      L     #Enc;
      T     #Data.Fall_Pos;
      L     #Data.Time_ms;
      T     #Data.Fall_ms;
      SET   ;
      S     #Data.Low;

S020: NOP   0;
NETWORK
TITLE =OFF Longer than Gap_Min = Real Gap - Close Packet

      A     #RUN;
      AN    #Sensor;
      A     #Data.Open;
      A     #Data.Low;
      JCN   S030;

      L     #Enc;
      L     #Data.Fall_Pos;
      -D    ;
      T     #D;
      L     L#0;
      >=D   ;
      JC    S031;

      L     #D;
      NEGD  ;
      T     #D;

S031: L     #D;
      L     #Gap_Min_Pulse;
      >=D   ;
      =     #CLOSE;

S030: NOP   0;
NETWORK
TITLE =Transfer End - Close Last Packet / Discard Covered One
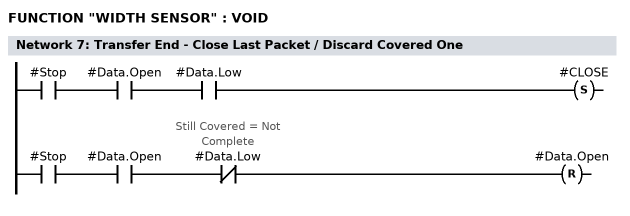

      A     #Stop;
      A     #Data.Open;
      A     #Data.Low;
      S     #CLOSE;
//;
      A     #Stop;
      A     #Data.Open;
      AN    #Data.Low; // Still Covered = Not Complete
      R     #Data.Open;

NETWORK
TITLE =Close Packet - Record Width

      A     #CLOSE;
      JCN   S090;

      A     #Data.Skip; // Partial Packet - Not Recorded
      JCN   S041;

      L     #Data.Skipped;
      L     1;
      +I    ;
      T     #Data.Skipped;
      JU    S049;

S041: L     #Data.Fall_Pos;
      L     #Data.Start_Pos;
      -D    ;
      T     #D;
      L     L#0;
      >=D   ;
      JC    S042;

      L     #D;
      NEGD  ;
      T     #D;

S042: L     #D;
      DTR   ;
      L     3.100000e-001;
      *R    ;
      RND   ;
      T     #MM;
      T     #Data.Last_Width_mm;
      L     #Data.Count;
      L     1;
      +I    ;
      T     #Data.Count;
      L     #MM;
      ITD   ;
      L     #Data.Width_Sum_mm;
      +D    ;
      T     #Data.Width_Sum_mm;
      L     #MM;
      L     #Data.Width_Min_mm;
      <I    ;
      JCN   S043;

      L     #MM;
      T     #Data.Width_Min_mm;

S043: L     #MM;
      L     #Data.Width_Max_mm;
      >I    ;
      JCN   S044;

      L     #MM;
      T     #Data.Width_Max_mm;

S044: L     #Data.Width_Sum_mm;
      L     #Data.Count;
      ITD   ;
      /D    ;
      T     #Data.Width_Avg_mm;
//;
      L     #Data.Fall_ms; // Width [mS] = Front -> End
      T     #Data.Last_Width_ms;
      L     #Data.Width_Sum_ms;
      +D    ;
      T     #Data.Width_Sum_ms;
      L     #Data.Count;
      ITD   ;
      /D    ;
      T     #Data.Width_Avg_ms;

S049: SET   ;
      R     #Data.Open;
      R     #Data.Low;
      R     #Data.Skip;

S090: NOP   0;
NETWORK
TITLE =Sensor State for Next Scan

      A     #Sensor;
      =     #Data.Was_On;
END_FUNCTION

FUNCTION "PACKET BLANKING" : VOID
TITLE =Packet Blanking - One Sensor (Shadow)
//v0.1 2026-11-19: one count per packet from a raw sensor, with the packet time
//measured at C10 (DB30 Width_ms_31, same speed on C11/C12/C21/C22).
//- Front (OFF->ON) counts if the belt has run >= Blank_Pct of a packet time
//  since the last count; an earlier front = sag of a U-Shape -> ignored.
//- Sensor still ON after Butt_Pct of a packet time = butted packet -> +1.
//- Time only runs while the belt runs (Run): a stop does not open the window.
//- Pulse: Pulse_ms long per counted packet (for FC8 later).
VERSION : 0.1


VAR_INPUT
  Sensor : BOOL ;	//Raw Packet Sensor
  Run : BOOL ;	//Belt Under the Sensor Runs
  Width_ms : INT ;	//Packet Time [mS]
  Blank_Pct : INT ;	//Blanking [%]
  Butt_Pct : INT ;	//Butted [%]
  Pulse_Len : INT ;	//Pulse [mS]
  Scan_mS : INT ;	//PLC Scan [mS]
END_VAR
VAR_OUTPUT
  Pulse : BOOL ;	//One Pulse per Counted Packet
END_VAR
VAR_IN_OUT
  D : "Blanking Struct";
END_VAR
VAR_TEMP
  BLANK : DINT ;
  BUTT : DINT ;
  CNT : BOOL ;
  BTD : BOOL ;
END_VAR
BEGIN
NETWORK
TITLE =Belt Run Time Since Last Count

      CLR   ;
      =     #CNT;
      =     #BTD;
//;
      A     #Run;
      JCN   B001;

      L     #D.T_ms;
      L     #Scan_mS;
      ITD   ;
      +D    ;
      T     #D.T_ms;
      L     #D.T_ms;
      L     L#60000;
      >D    ; // Clamp 60s
      JCN   B001;

      L     L#60000;
      T     #D.T_ms;

B001: NOP   0;
NETWORK
TITLE =Windows [mS]

      L     #Width_ms;
      ITD   ;
      L     #Blank_Pct;
      ITD   ;
      *D    ;
      L     L#100;
      /D    ;
      T     #BLANK;
//;
      L     #Width_ms;
      ITD   ;
      L     #Butt_Pct;
      ITD   ;
      *D    ;
      L     L#100;
      /D    ;
      T     #BUTT;
NETWORK
TITLE =Front - Count, or Ignore Inside Blanking (Sag)

      A     #Sensor;
      AN    #D.Was_On;
      JCN   B010;

      L     #D.Raw;
      L     1;
      +I    ;
      T     #D.Raw;
//;
      L     #D.T_ms;
      L     #BLANK;
      >=D   ;
      =     #CNT; // Front Counts
      JC    B010;

      L     #D.Sag; // Front Inside Blanking = Sag
      L     1;
      +I    ;
      T     #D.Sag;

B010: NOP   0;
NETWORK
TITLE =Sensor Still ON - Butted Packet

      A     #Sensor;
      A     #Run;
      AN    #CNT;
      JCN   B020;

      L     #D.T_ms;
      L     #BUTT;
      >=D   ;
      JCN   B020;

      L     #D.Butt;
      L     1;
      +I    ;
      T     #D.Butt;
      SET   ;
      =     #CNT;
      =     #BTD; // Next Butted Packet One Packet Time Later

B020: NOP   0;
NETWORK
TITLE =Count + Pulse

      A     #CNT;
      JCN   B030;

      L     #D.Count;
      L     1;
      +I    ;
      T     #D.Count;
      L     L#0;
      T     #D.T_ms;
      A     #BTD;
      JCN   B032;

      L     #BUTT; // Butted: T = Butt - Packet Time
      L     #Width_ms;
      ITD   ;
      -D    ;
      T     #D.T_ms;

B032: L     #Pulse_Len;
      T     #D.Pulse_ms;

B030: L     #D.Pulse_ms;
      L     0;
      >I    ;
      =     #Pulse;
      =     #D.Pulse;
      JCN   B031;

      L     #D.Pulse_ms;
      L     #Scan_mS;
      -I    ;
      T     #D.Pulse_ms;

B031: A     #Sensor;
      =     #D.Was_On;
END_FUNCTION

FUNCTION "PACKET POSITIONING" : VOID
TITLE =Packet Positioning - Flipper C7 + Pusher 2 C9 - Stop Time per Lengt
//v1.0 2026-11-23: called by FC942 v1.0. Picks the stop time of the length class
//of the packets (C4 measurement), lights the class lamp, and lets the operator
//change that class time with the HMI arrows (+/- Step_ms, Min_ms...Max_ms).
//Writes only DB15 "PACKET POSITION DB". Empty table = Default_ms = 1.5 s as before.
//v1.1 2026-11-24: HMI packet drawing: length (DBW86) + width class bits (DBX90.x).
//v1.2 2026-11-24: renumbered FC1221 -> FC1215 (same name "FLIPPER POS ADJ", no
//code change). FC942 calls it by name.
//v1.3 2026-11-24: renamed "PACKET POSITIONING". + C9 Pusher 2 conveyor: same
//length class, own table / arrows, default = "HMI_DB".CONV_9_POS_mS x 10 (as
//before). Output C9_Stop_S5T for FC950 v1.0 Timer 62.
//v1.4 2026-11-24: C9 HMI drawing: C9_Pos_Bits (one of 16 lateral positions).
//v1.5 2026-11-24: DB15 symbol renamed "PACKET POSITION DB" - no code change.
VERSION : 1.5


VAR_TEMP
  CLASS : INT ;
  T_TAB : INT ;
  T_NEW : INT ;
  T_DEF : INT ;
  T_TIME : TIME ;
  S5 : S5TIME ;
END_VAR
BEGIN
NETWORK
TITLE =Packet Length -> Class (15 mm Steps from 510 mm, 0...31)

      L     "HOUSE_KEEPING DB".C4_Packet_Length_mm;
      T     "PACKET POSITION DB".Length_mm;
      L     510;
      -I    ;
      L     15;
      /I    ;
      T     #CLASS;
      L     0;
      >=I   ;
      JC    K001;

      L     0;
      T     #CLASS;

K001: L     #CLASS;
      L     31;
      <=I   ;
      JC    K002;

      L     31;
      T     #CLASS;

K002: L     #CLASS;
      T     "PACKET POSITION DB".Class;
//;
      L     #CLASS; // Class Lamp: Bit = Class
      L     L#1;
      SLD   ;
      T     "PACKET POSITION DB".Class_Lamps;
NETWORK
TITLE =C7 Flipper - Read the Class Time (Time_ms[Class], DB15.DBW22 + 2 x

      L     #CLASS;
      SLW   1;
      L     22;
      +I    ;
      SLD   3;
      LAR1  ;
      OPN   "PACKET POSITION DB";
      L     DBW [AR1,P#0.0];
      T     #T_TAB;
NETWORK
TITLE =C7 Flipper - HMI Arrows / Reset - Change This Class Time
//The HMI sets Plus_PB / Minus_PB / Reset_PB, the PLC resets them after use:
//one press = one step.
      L     #T_TAB; // Start From the Time Used (0 = Default)
      L     0;
      <>I   ;
      JC    K010;

      L     "PACKET POSITION DB".Default_ms;
      JU    K011;

K010: L     #T_TAB;
K011: T     #T_NEW;
//;
      A     "PACKET POSITION DB".Plus_PB;
      JCN   K012;

      L     #T_NEW;
      L     "PACKET POSITION DB".Step_ms;
      +I    ;
      T     #T_NEW;

K012: A     "PACKET POSITION DB".Minus_PB;
      JCN   K013;

      L     #T_NEW;
      L     "PACKET POSITION DB".Step_ms;
      -I    ;
      T     #T_NEW;

K013: L     #T_NEW; // Clamp Min...Max
      L     "PACKET POSITION DB".Min_ms;
      >=I   ;
      JC    K014;

      L     "PACKET POSITION DB".Min_ms;
      T     #T_NEW;

K014: L     #T_NEW;
      L     "PACKET POSITION DB".Max_ms;
      <=I   ;
      JC    K015;

      L     "PACKET POSITION DB".Max_ms;
      T     #T_NEW;

K015: NOP   0;
NETWORK
TITLE =C7 Flipper - Write Back After an Arrow / Reset

      A     "PACKET POSITION DB".Reset_PB;
      JCN   K020;

      L     0; // Class Back to Default
      T     #T_TAB;
      JU    K021;

K020: A(    ;
      O     "PACKET POSITION DB".Plus_PB;
      O     "PACKET POSITION DB".Minus_PB;
      )     ;
      JCN   K022;

      L     #T_NEW;
      T     #T_TAB;

K021: L     #CLASS;
      SLW   1;
      L     22;
      +I    ;
      SLD   3;
      LAR1  ;
      OPN   "PACKET POSITION DB";
      L     #T_TAB;
      T     DBW [AR1,P#0.0];

K022: SET   ; // Momentary: Reset by the PLC
      R     "PACKET POSITION DB".Plus_PB;
      R     "PACKET POSITION DB".Minus_PB;
      R     "PACKET POSITION DB".Reset_PB;
NETWORK
TITLE =HMI Packet Drawing - Length + Width Class (4 Pairs of Level Meters)
//Width = C10 measured width (DB30 Width_mm_Cal, last verified, same order).
//0 (not measured yet) = smallest class.
      L     "PACKET POSITION DB".Length_mm;
      T     "PACKET POSITION DB".Disp_Length_mm;
//;
      L     "PACKET WIDTH DB".Width_mm_Cal;
      T     "PACKET POSITION DB".Width_mm;
//;
      L     "PACKET POSITION DB".Width_mm;
      L     "PACKET POSITION DB".Width_Lim_1;
      <I    ;
      =     "PACKET POSITION DB".Width_Class_1;
//;
      A(    ;
      L     "PACKET POSITION DB".Width_mm;
      L     "PACKET POSITION DB".Width_Lim_1;
      >=I   ;
      )     ;
      A(    ;
      L     "PACKET POSITION DB".Width_mm;
      L     "PACKET POSITION DB".Width_Lim_2;
      <I    ;
      )     ;
      =     "PACKET POSITION DB".Width_Class_2;
//;
      A(    ;
      L     "PACKET POSITION DB".Width_mm;
      L     "PACKET POSITION DB".Width_Lim_2;
      >=I   ;
      )     ;
      A(    ;
      L     "PACKET POSITION DB".Width_mm;
      L     "PACKET POSITION DB".Width_Lim_3;
      <I    ;
      )     ;
      =     "PACKET POSITION DB".Width_Class_3;
//;
      L     "PACKET POSITION DB".Width_mm;
      L     "PACKET POSITION DB".Width_Lim_3;
      >=I   ;
      =     "PACKET POSITION DB".Width_Class_4;
NETWORK
TITLE =C7 Flipper - Stop Time Used -> S5TIME for FC942 Timer 42

      L     #T_TAB;
      L     0;
      <>I   ;
      A     "PACKET POSITION DB".Use_Table;
      JC    K030;

      L     "PACKET POSITION DB".Default_ms;
      JU    K031;

K030: L     #T_TAB;
K031: T     "PACKET POSITION DB".Time_Used_ms;
      ITD   ;
      T     #T_TIME;

      CALL "TIM_S5TI" (
           IN                       := #T_TIME,
           RET_VAL                  := #S5);

      L     #S5;
      T     "PACKET POSITION DB".Stop_S5T;
NETWORK
TITLE =C9 Pusher 2 - Read the Class Time (C9_Time_ms[Class], DB15.DBW108 +

      L     "PACKET POSITION DB".Class;
      T     #CLASS;
      SLW   1;
      L     108;
      +I    ;
      SLD   3;
      LAR1  ;
      OPN   "PACKET POSITION DB";
      L     DBW [AR1,P#0.0];
      T     #T_TAB;
//;
      L     "HMI_DB".CONV_9_POS_mS; // C9 Default = HMI Time x 10 mS (as Before)
      L     10;
      *I    ;
      T     #T_DEF;
NETWORK
TITLE =C9 Pusher 2 - HMI Arrows / Reset - Change This Class Time

      L     #T_TAB;
      L     0;
      <>I   ;
      JC    C010;

      L     #T_DEF;
      JU    C011;

C010: L     #T_TAB;
C011: T     #T_NEW;
//;
      A     "PACKET POSITION DB".C9_Plus_PB;
      JCN   C012;

      L     #T_NEW;
      L     "PACKET POSITION DB".Step_ms;
      +I    ;
      T     #T_NEW;

C012: A     "PACKET POSITION DB".C9_Minus_PB;
      JCN   C013;

      L     #T_NEW;
      L     "PACKET POSITION DB".Step_ms;
      -I    ;
      T     #T_NEW;

C013: L     #T_NEW; // Clamp 1...Max (0 Means Default)
      L     1;
      >=I   ;
      JC    C014;

      L     1;
      T     #T_NEW;

C014: L     #T_NEW;
      L     "PACKET POSITION DB".Max_ms;
      <=I   ;
      JC    C015;

      L     "PACKET POSITION DB".Max_ms;
      T     #T_NEW;

C015: NOP   0;
NETWORK
TITLE =C9 Pusher 2 - Write Back After an Arrow / Reset

      A     "PACKET POSITION DB".C9_Reset_PB;
      JCN   C020;

      L     0; // Class Back to Default
      T     #T_TAB;
      JU    C021;

C020: A(    ;
      O     "PACKET POSITION DB".C9_Plus_PB;
      O     "PACKET POSITION DB".C9_Minus_PB;
      )     ;
      JCN   C022;

      L     #T_NEW;
      T     #T_TAB;

C021: L     #CLASS;
      SLW   1;
      L     108;
      +I    ;
      SLD   3;
      LAR1  ;
      OPN   "PACKET POSITION DB";
      L     #T_TAB;
      T     DBW [AR1,P#0.0];

C022: SET   ; // Momentary: Reset by the PLC
      R     "PACKET POSITION DB".C9_Plus_PB;
      R     "PACKET POSITION DB".C9_Minus_PB;
      R     "PACKET POSITION DB".C9_Reset_PB;
NETWORK
TITLE =C9 Pusher 2 - Stop Time Used -> S5TIME for FC950 Timer 62

      L     #T_TAB;
      L     0;
      <>I   ;
      A     "PACKET POSITION DB".C9_Use_Table;
      JC    C030;

      L     #T_DEF;
      JU    C031;

C030: L     #T_TAB;
C031: T     "PACKET POSITION DB".C9_Time_Used_ms;
      ITD   ;
      T     #T_TIME;

      CALL "TIM_S5TI" (
           IN                       := #T_TIME,
           RET_VAL                  := #S5);

      L     #S5;
      T     "PACKET POSITION DB".C9_Stop_S5T;
NETWORK
TITLE =C9 Pusher 2 - HMI Drawing: 1 of 16 Lateral Positions (Longer Time =

      L     "PACKET POSITION DB".C9_View_Step_ms; // Step 0 -> Copy 0
      L     0;
      >I    ;
      JC    C040;

      L     0;
      JU    C042;

C040: L     "PACKET POSITION DB".C9_Time_Used_ms;
      L     "PACKET POSITION DB".C9_View_Min_ms;
      -I    ;
      L     "PACKET POSITION DB".C9_View_Step_ms;
      /I    ;
      T     #T_NEW;
      L     0;
      >=I   ;
      JC    C041;

      L     0;
      T     #T_NEW;

C041: L     #T_NEW;
      L     15;
      <=I   ;
      L     #T_NEW;
      JC    C042;

      L     15;
C042: T     "PACKET POSITION DB".C9_Pos_Step;
//;
      L     "PACKET POSITION DB".C9_Pos_Step; // One Bit = Step
      L     L#1;
      SLD   ;
      T     "PACKET POSITION DB".C9_Pos_Bits;
END_FUNCTION

FUNCTION "LAUER CALL" : VOID
TITLE =Lauer Call
// TEXT ORG
NAME : TEXTORG
VERSION : 0.0

BEGIN
NETWORK
TITLE =

      OPN   "DB LAUER";

NETWORK
TITLE =Reset & Preset
//When the communication/control byte is in a neutral state, and those two
//internal flags are off, the FC restores default preset values in the Lauer DB.
      A(    ;
      L     "MB 150";
      L     W#16#FFF7;
      AW    ;
      L     W#16#0;
      )     ;
      ==I   ;
      AN    "M 151.6";
      AN    "M 151.7";
      JC    M001;
      JU    M002;

M001: L     2#0;
      T     DBW   76;
//;
      L     2#111100000000;
      T     DBW   72;
//;
      L     2#11100000000001;
      T     DBW   74;
//;
      L     W#16#0;
      T     DBW   32;

M002: NOP   0;
NETWORK
TITLE =
//transfer keypad/page/request words
//avoid repeated copying every scan
//only copy
//once per trigger edge/state
      A     "M 0.3";
      AN    "M 200.0";
      JC    M003;
      A     "M 0.2";
      AN    "M 200.1";
      JC    M004;
      JU    M005;

M003: L     "MW 150";
      T     "MW 118";
//;
      L     "MW 152";
      T     "MW 120";
//;
      A     "M 0.3";
      S     "M 200.0";
      R     "M 200.1";
      JU    M005;

M004: L     "MW 118";
      T     "MW 150";
//;
      L     "MW 120";
      T     "MW 152";
//;
      A     "M 0.2";
      S     "M 200.1";
      R     "M 200.0";

M005: NOP   0;
NETWORK
TITLE =
//reopen "DB LAUER"
//
//load DBW48
//
//call LAUER KEYS 1
      OPN   "DB LAUER";
      L     DBW   48;
      CALL "LAUER KEYS 1" ;
NETWORK
TITLE =

      CALL "LAUER SERVICE" ;

NETWORK
TITLE =

      CALL "LAUER KEYS 2" ;

NETWORK
TITLE =

      CALL "LAUER KEYS 3" ;

NETWORK
TITLE =

      CALL "LAUER MESSAGE1" ;

NETWORK
TITLE =

//      CALL  "LAUER"

NETWORK
TITLE =

      CALL "LAUER MESSAGE2" ;

END_FUNCTION

FUNCTION "SETUP" : VOID
TITLE =Setup Values
//Do Not Change These Values !!!
NAME : SETUP
VERSION : 0.1

BEGIN
NETWORK
TITLE =Setup Values - Slat Conveyor 3

      L     8000;
      T     "COLLATORS DB".Conveyor_Length_C3;
NETWORK
TITLE =Setup Values - Conveyor 4

      L     800; //900
      T     "COLLATORS DB".Surface_Length_C4;
NETWORK
TITLE =Setup Value  - TurnTable - Need " Packet IN " to Start

      S     "M 47.4";

NETWORK
TITLE =Setup Values - Conveyor 10

      L     13000;
      T     "COLLATORS DB".Surface_Length_10;
NETWORK
TITLE =Counter Setup


      S     "M 167.7";
NETWORK
TITLE =Packet Counter Constants 11.0 & 5.5

      L     1.000000e+001;
      T     "DB UTILITY".LENGTH_CONST;
//;
      L     5.200000e-001;
      T     "DB UTILITY".WIDTH_CONST;
NETWORK
TITLE =HMI - Conveyor Time

      L     150;
      T     "HMI_DB".CONV_7_POS_mS;
//;
      L     30;
      T     "HMI_DB".CONV_8_POS_FWD_mS;
//;
      L     70;
      T     "HMI_DB".CONV_8_POS_REV_mS;
//;
      L     15;
      T     "HMI_DB".CONV_9_POS_mS;
NETWORK
TITLE =HMI Control - Reset

      R     "HMI_DB".SERVICE_SW_1_STATUS;
      R     "HMI_DB".SERVICE_SW_2_STATUS;
      R     "HMI_DB".SERVICE_SW_3_STATUS;
      R     "HMI_DB".SERVICE_SW_1_2_STATUS;
END_FUNCTION

FUNCTION "SENSOR DE-BOUNCER" : VOID
TITLE =Sensor Debouncer
//Counting Foul Sensor Switching of less than PreSet Time
VERSION : 0.2


VAR_INPUT
  Bit_0 : BOOL ;
  Bit_1 : BOOL ;
  Preset_mS : INT ;
  Debounce_mS : INT ;
  Plc_Scan_mS : INT ;
END_VAR
VAR_IN_OUT
  Rising_Pulse_1 : BOOL ;	//Db Struct
  Rising_Pulse_2 : BOOL ;	//Db Struct
  Rising_Pulse_3 : BOOL ;	//Db Struct
  Rising_Pulse_4 : BOOL ;	//Db Struct
  Rising_Pulse_5 : BOOL ;	//Db Struct
  Rising_Pulse_6 : BOOL ;	//Db Struct
  Rising_Pulse_7 : BOOL ;	//Db Struct
  Rising_Pulse_8 : BOOL ;	//Db Struct
  Memory_Bit_1 : BOOL ;	//Db Struct
  Memory_Bit_2 : BOOL ;	//Db Struct
  Memory_Bit_3 : BOOL ;	//Db Struct
  Memory_Bit_4 : BOOL ;	//Db Struct
  Memory_Bit_5 : BOOL ;	//Db Struct
  Memory_Bit_6 : BOOL ;	//Db Struct
  Spare_1 : BOOL ;	//Db Struct
  Spare_2 : BOOL ;	//Db Struct
  Word_Buffer_1 : INT ;	//Db Struct
  Word_Buffer_2 : INT ;	//Db Struct
  Word_Result : INT ;	//Db Struct
  Word_Count_Limit : INT ;	//Db Data
  Word_Count : INT ;	//Db/HMI Data
END_VAR
VAR_TEMP
  MEMORY_1 : BOOL ;
  MEMORY_2 : BOOL ;
  MEMORY_3 : BOOL ;
END_VAR
BEGIN
NETWORK
TITLE =Init on First Call

      A     #Memory_Bit_6;
      JNB   INI1;
      JU    INI2;

INI1: L     0;
      T     #Word_Buffer_1;
      T     #Word_Buffer_2;
      R     #Memory_Bit_1;
      R     #Memory_Bit_2;
      R     #Memory_Bit_3;
      R     #Memory_Bit_4;
      R     #Memory_Bit_5;
      S     #Memory_Bit_6;

INI2: NOP   0;

NETWORK
TITLE =Input Bits - Start Event
//- #Bit_0 : Conveyor X InFeed Sensor
//- #Bit_1 : Conveyor X Exit Sensor
      A     #Bit_0;
      FP    #Rising_Pulse_1;
      JNB   K001;
      L     0;
      T     #Word_Buffer_1;
      R     #Memory_Bit_4;
      S     #Memory_Bit_1;

K001: NOP   0;

      A     #Bit_1;
      FP    #Rising_Pulse_2;
      JNB   K002;
      L     0;
      T     #Word_Buffer_2;
      S     #Memory_Bit_2;

K002: NOP   0;

NETWORK
TITLE =TimeBase
//TimeBase -> ScanTime
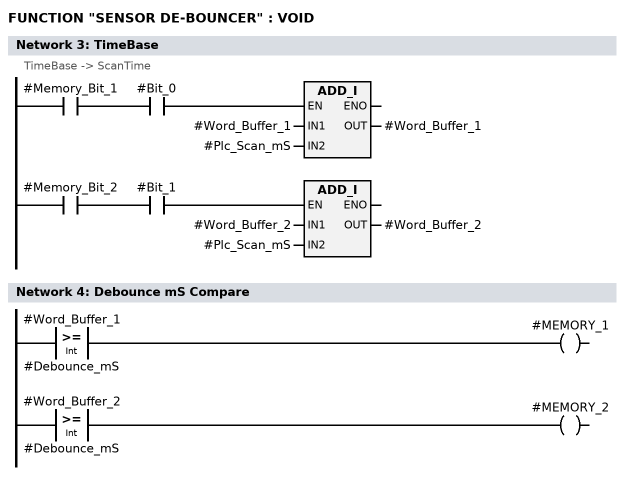
      A     #Memory_Bit_1;
      A     #Bit_0;
      JNB   K003;
      L     #Word_Buffer_1;
      L     #Plc_Scan_mS;
      +I    ;
      T     #Word_Buffer_1;

K003: NOP   0;

      A     #Memory_Bit_2;
      A     #Bit_1;
      JNB   K004;
      L     #Word_Buffer_2;
      L     #Plc_Scan_mS;
      +I    ;
      T     #Word_Buffer_2;

K004: NOP   0;

NETWORK
TITLE =Debounce mS Compare

      A(    ;
      L     #Word_Buffer_1;
      L     #Debounce_mS;
      >=I   ;
      )     ;
      =     #MEMORY_1;
//;
      A(    ;
      L     #Word_Buffer_2;
      L     #Debounce_mS;
      >=I   ;
      )     ;
      =     #MEMORY_2;

NETWORK
TITLE =Add to Packet Number with Bit_0
//Validated ON event on Bit_0 adds +1 one time
      A     #Memory_Bit_1;
      A     #MEMORY_1;
      A     #Bit_0;
      FP    #Rising_Pulse_4;
      JNB   K005;
      L     #Word_Count;
      L     1;
      +I    ;
      T     #Word_Count;
      R     #Memory_Bit_1;

K005: NOP   0;

NETWORK
TITLE =Subtract from Packet Number with Bit_1
//Validated ON event on Bit_1 subtracts -1 on falling edge
      AN    #Bit_1;
      FP    #Rising_Pulse_5;
      JNB   K006;

      A     #Memory_Bit_2;
      A     #MEMORY_2;
      JNB   K006;
//;
      L     #Word_Count;
      L     1;
      -I    ;
      T     #Word_Count;
      R     #Memory_Bit_2;

K006: NOP   0;

NETWORK
TITLE =Clamp Packet Number
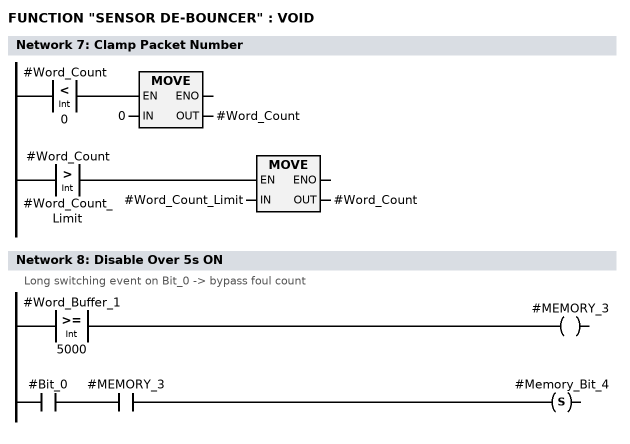

      L     #Word_Count;
      L     0;
      <I    ;
      JNB   K007;
      L     0;
      T     #Word_Count;

K007: NOP   0;

      L     #Word_Count;
      L     #Word_Count_Limit;
      >I    ;
      JNB   K008;
      L     #Word_Count_Limit;
      T     #Word_Count;

K008: NOP   0;

NETWORK
TITLE =Disable Over 5s ON
//Long switching event on Bit_0 -> bypass foul count
      L     #Word_Buffer_1;
      L     5000;
      >=I   ;
      =     #MEMORY_3;
//;
      A     #Bit_0;
      A     #MEMORY_3;
      S     #Memory_Bit_4;

NETWORK
TITLE =Result
//Word_Result +1 if Bit_0 turns OFF before Preset_mS and was not bypassed
      AN    #Bit_0;
      FP    #Rising_Pulse_6;
      JNB   K009;

      A     #Memory_Bit_1;
      AN    #Memory_Bit_4;
      JNB   K010;
//;
      L     #Word_Buffer_1;
      L     #Preset_mS;
      <I    ;
      JNB   K010;
//;
      L     #Word_Result;
      L     1;
      +I    ;
      T     #Word_Result;

K010: R     #Memory_Bit_1;
      R     #Memory_Bit_4;
      L     0;
      T     #Word_Buffer_1;

K009: NOP   0;

NETWORK
TITLE =Reset Exit Event on Falling Edge

      AN    #Bit_1;
      FP    #Rising_Pulse_7;
      JNB   K011;
      R     #Memory_Bit_2;
      L     0;
      T     #Word_Buffer_2;

K011: NOP   0;

END_FUNCTION

FUNCTION "SENSOR CHECK CALLS" : VOID
TITLE =
VERSION : 0.1

BEGIN
NETWORK
TITLE =
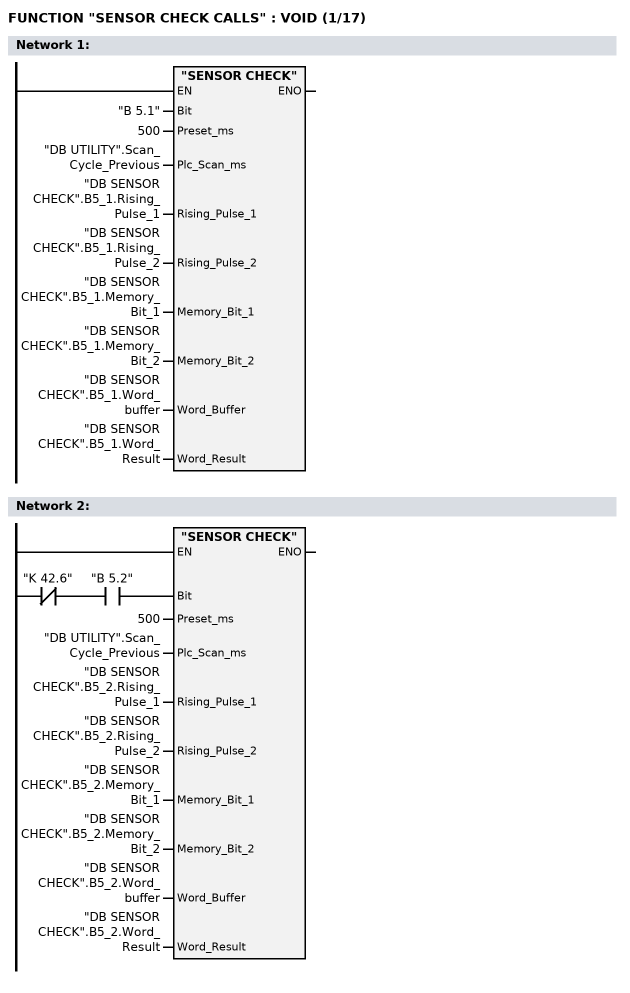

      CALL "SENSOR CHECK" (
           Bit                      := "B 5.1",
           Preset_ms                := 500,
           Plc_Scan_ms              := "DB UTILITY".Scan_Cycle_Previous,
           Rising_Pulse_1           := "DB SENSOR CHECK".B5_1.Rising_Pulse_1,
           Rising_Pulse_2           := "DB SENSOR CHECK".B5_1.Rising_Pulse_2,
           Memory_Bit_1             := "DB SENSOR CHECK".B5_1.Memory_Bit_1,
           Memory_Bit_2             := "DB SENSOR CHECK".B5_1.Memory_Bit_2,
           Word_Buffer              := "DB SENSOR CHECK".B5_1.Word_buffer,
           Word_Result              := "DB SENSOR CHECK".B5_1.Word_Result);

NETWORK
TITLE =

      AN    "K 42.6";
      A     "B 5.2";
      =     L      0.0;
//;
      CALL "SENSOR CHECK" (
           Bit                      := L      0.0,
           Preset_ms                := 500,
           Plc_Scan_ms              := "DB UTILITY".Scan_Cycle_Previous,
           Rising_Pulse_1           := "DB SENSOR CHECK".B5_2.Rising_Pulse_1,
           Rising_Pulse_2           := "DB SENSOR CHECK".B5_2.Rising_Pulse_2,
           Memory_Bit_1             := "DB SENSOR CHECK".B5_2.Memory_Bit_1,
           Memory_Bit_2             := "DB SENSOR CHECK".B5_2.Memory_Bit_2,
           Word_Buffer              := "DB SENSOR CHECK".B5_2.Word_buffer,
           Word_Result              := "DB SENSOR CHECK".B5_2.Word_Result);

NETWORK
TITLE =
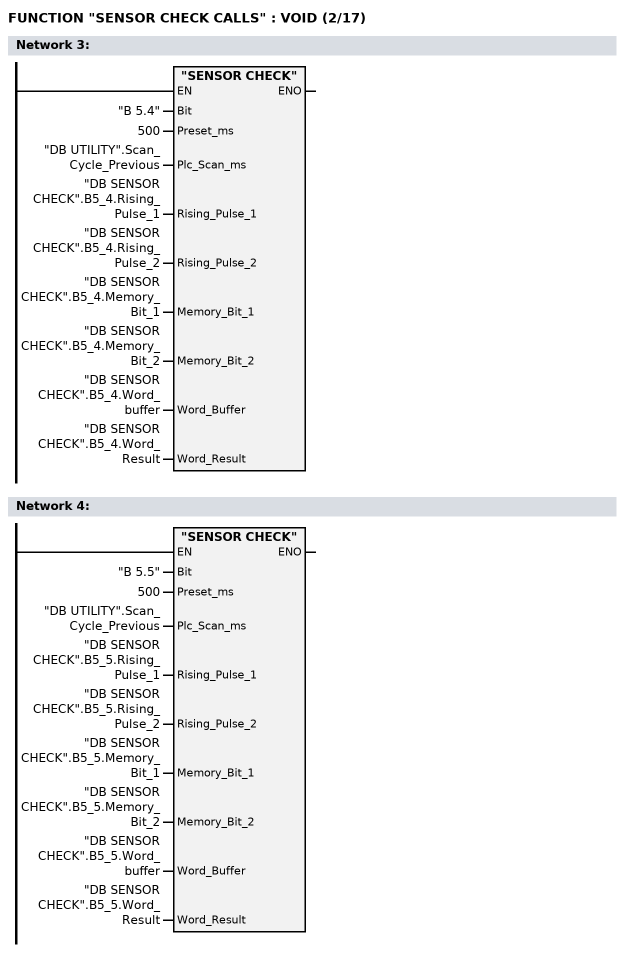

      CALL "SENSOR CHECK" (
           Bit                      := "B 5.4",
           Preset_ms                := 500,
           Plc_Scan_ms              := "DB UTILITY".Scan_Cycle_Previous,
           Rising_Pulse_1           := "DB SENSOR CHECK".B5_4.Rising_Pulse_1,
           Rising_Pulse_2           := "DB SENSOR CHECK".B5_4.Rising_Pulse_2,
           Memory_Bit_1             := "DB SENSOR CHECK".B5_4.Memory_Bit_1,
           Memory_Bit_2             := "DB SENSOR CHECK".B5_4.Memory_Bit_2,
           Word_Buffer              := "DB SENSOR CHECK".B5_4.Word_buffer,
           Word_Result              := "DB SENSOR CHECK".B5_4.Word_Result);

NETWORK
TITLE =

      CALL "SENSOR CHECK" (
           Bit                      := "B 5.5",
           Preset_ms                := 500,
           Plc_Scan_ms              := "DB UTILITY".Scan_Cycle_Previous,
           Rising_Pulse_1           := "DB SENSOR CHECK".B5_5.Rising_Pulse_1,
           Rising_Pulse_2           := "DB SENSOR CHECK".B5_5.Rising_Pulse_2,
           Memory_Bit_1             := "DB SENSOR CHECK".B5_5.Memory_Bit_1,
           Memory_Bit_2             := "DB SENSOR CHECK".B5_5.Memory_Bit_2,
           Word_Buffer              := "DB SENSOR CHECK".B5_5.Word_buffer,
           Word_Result              := "DB SENSOR CHECK".B5_5.Word_Result);

NETWORK
TITLE =
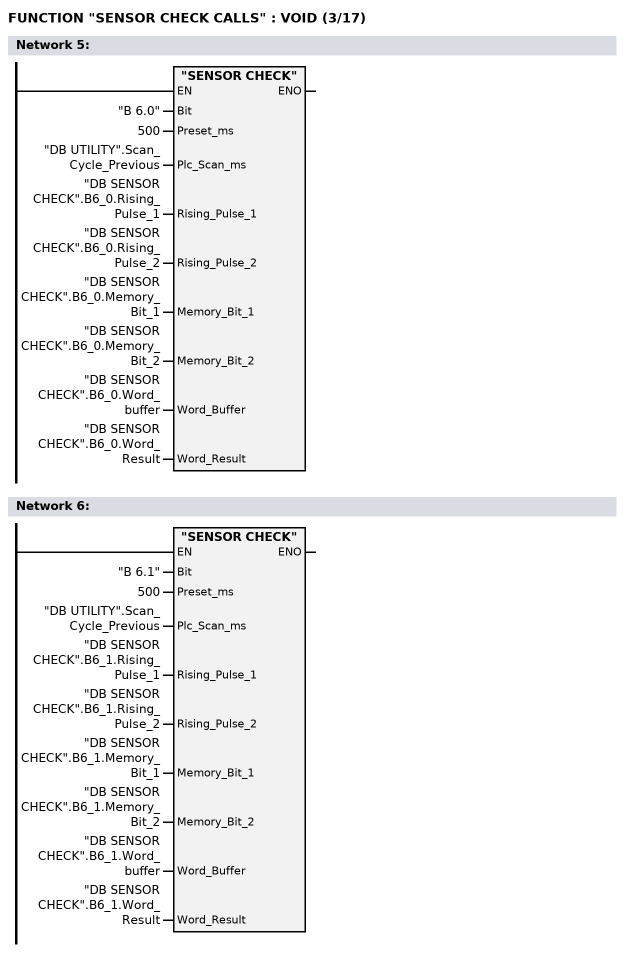

      CALL "SENSOR CHECK" (
           Bit                      := "B 6.0",
           Preset_ms                := 500,
           Plc_Scan_ms              := "DB UTILITY".Scan_Cycle_Previous,
           Rising_Pulse_1           := "DB SENSOR CHECK".B6_0.Rising_Pulse_1,
           Rising_Pulse_2           := "DB SENSOR CHECK".B6_0.Rising_Pulse_2,
           Memory_Bit_1             := "DB SENSOR CHECK".B6_0.Memory_Bit_1,
           Memory_Bit_2             := "DB SENSOR CHECK".B6_0.Memory_Bit_2,
           Word_Buffer              := "DB SENSOR CHECK".B6_0.Word_buffer,
           Word_Result              := "DB SENSOR CHECK".B6_0.Word_Result);

NETWORK
TITLE =

      CALL "SENSOR CHECK" (
           Bit                      := "B 6.1",
           Preset_ms                := 500,
           Plc_Scan_ms              := "DB UTILITY".Scan_Cycle_Previous,
           Rising_Pulse_1           := "DB SENSOR CHECK".B6_1.Rising_Pulse_1,
           Rising_Pulse_2           := "DB SENSOR CHECK".B6_1.Rising_Pulse_2,
           Memory_Bit_1             := "DB SENSOR CHECK".B6_1.Memory_Bit_1,
           Memory_Bit_2             := "DB SENSOR CHECK".B6_1.Memory_Bit_2,
           Word_Buffer              := "DB SENSOR CHECK".B6_1.Word_buffer,
           Word_Result              := "DB SENSOR CHECK".B6_1.Word_Result);

NETWORK
TITLE =
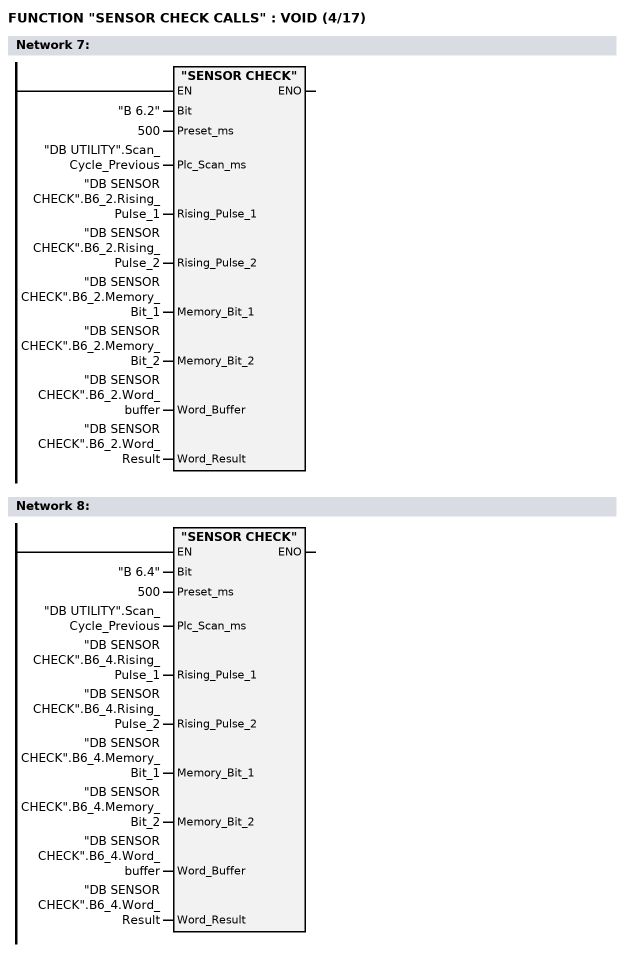

      CALL "SENSOR CHECK" (
           Bit                      := "B 6.2",
           Preset_ms                := 500,
           Plc_Scan_ms              := "DB UTILITY".Scan_Cycle_Previous,
           Rising_Pulse_1           := "DB SENSOR CHECK".B6_2.Rising_Pulse_1,
           Rising_Pulse_2           := "DB SENSOR CHECK".B6_2.Rising_Pulse_2,
           Memory_Bit_1             := "DB SENSOR CHECK".B6_2.Memory_Bit_1,
           Memory_Bit_2             := "DB SENSOR CHECK".B6_2.Memory_Bit_2,
           Word_Buffer              := "DB SENSOR CHECK".B6_2.Word_buffer,
           Word_Result              := "DB SENSOR CHECK".B6_2.Word_Result);

NETWORK
TITLE =

      CALL "SENSOR CHECK" (
           Bit                      := "B 6.4",
           Preset_ms                := 500,
           Plc_Scan_ms              := "DB UTILITY".Scan_Cycle_Previous,
           Rising_Pulse_1           := "DB SENSOR CHECK".B6_4.Rising_Pulse_1,
           Rising_Pulse_2           := "DB SENSOR CHECK".B6_4.Rising_Pulse_2,
           Memory_Bit_1             := "DB SENSOR CHECK".B6_4.Memory_Bit_1,
           Memory_Bit_2             := "DB SENSOR CHECK".B6_4.Memory_Bit_2,
           Word_Buffer              := "DB SENSOR CHECK".B6_4.Word_buffer,
           Word_Result              := "DB SENSOR CHECK".B6_4.Word_Result);

NETWORK
TITLE =
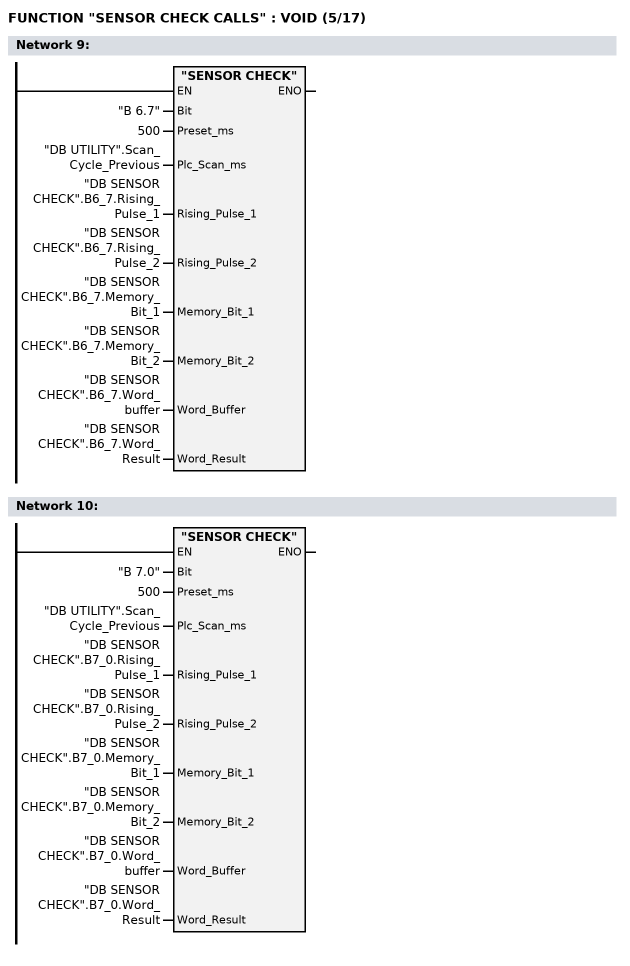

      CALL "SENSOR CHECK" (
           Bit                      := "B 6.7",
           Preset_ms                := 500,
           Plc_Scan_ms              := "DB UTILITY".Scan_Cycle_Previous,
           Rising_Pulse_1           := "DB SENSOR CHECK".B6_7.Rising_Pulse_1,
           Rising_Pulse_2           := "DB SENSOR CHECK".B6_7.Rising_Pulse_2,
           Memory_Bit_1             := "DB SENSOR CHECK".B6_7.Memory_Bit_1,
           Memory_Bit_2             := "DB SENSOR CHECK".B6_7.Memory_Bit_2,
           Word_Buffer              := "DB SENSOR CHECK".B6_7.Word_buffer,
           Word_Result              := "DB SENSOR CHECK".B6_7.Word_Result);

NETWORK
TITLE =

      CALL "SENSOR CHECK" (
           Bit                      := "B 7.0",
           Preset_ms                := 500,
           Plc_Scan_ms              := "DB UTILITY".Scan_Cycle_Previous,
           Rising_Pulse_1           := "DB SENSOR CHECK".B7_0.Rising_Pulse_1,
           Rising_Pulse_2           := "DB SENSOR CHECK".B7_0.Rising_Pulse_2,
           Memory_Bit_1             := "DB SENSOR CHECK".B7_0.Memory_Bit_1,
           Memory_Bit_2             := "DB SENSOR CHECK".B7_0.Memory_Bit_2,
           Word_Buffer              := "DB SENSOR CHECK".B7_0.Word_buffer,
           Word_Result              := "DB SENSOR CHECK".B7_0.Word_Result);

NETWORK
TITLE =
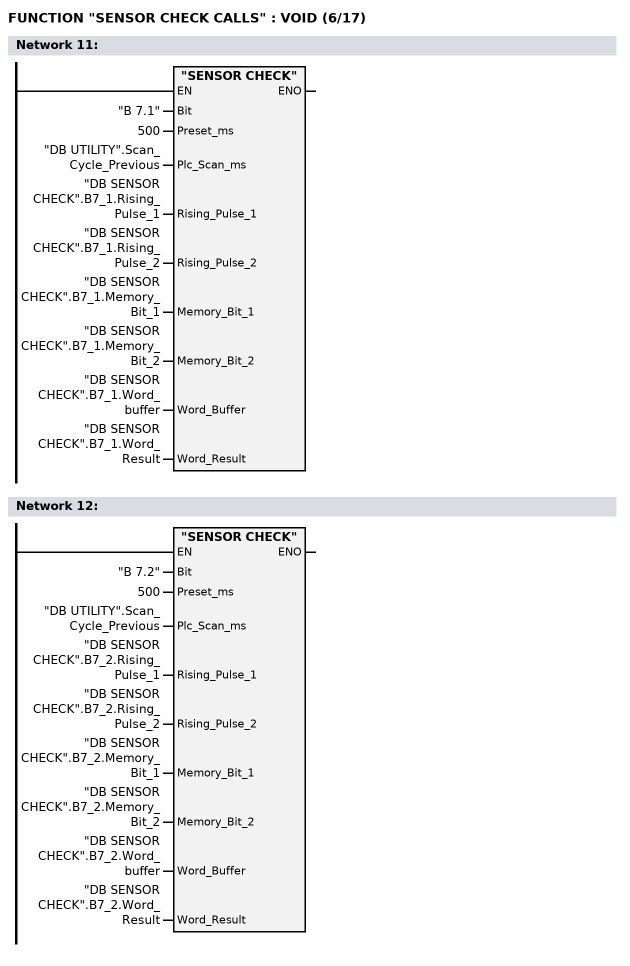

      CALL "SENSOR CHECK" (
           Bit                      := "B 7.1",
           Preset_ms                := 500,
           Plc_Scan_ms              := "DB UTILITY".Scan_Cycle_Previous,
           Rising_Pulse_1           := "DB SENSOR CHECK".B7_1.Rising_Pulse_1,
           Rising_Pulse_2           := "DB SENSOR CHECK".B7_1.Rising_Pulse_2,
           Memory_Bit_1             := "DB SENSOR CHECK".B7_1.Memory_Bit_1,
           Memory_Bit_2             := "DB SENSOR CHECK".B7_1.Memory_Bit_2,
           Word_Buffer              := "DB SENSOR CHECK".B7_1.Word_buffer,
           Word_Result              := "DB SENSOR CHECK".B7_1.Word_Result);

NETWORK
TITLE =

      CALL "SENSOR CHECK" (
           Bit                      := "B 7.2",
           Preset_ms                := 500,
           Plc_Scan_ms              := "DB UTILITY".Scan_Cycle_Previous,
           Rising_Pulse_1           := "DB SENSOR CHECK".B7_2.Rising_Pulse_1,
           Rising_Pulse_2           := "DB SENSOR CHECK".B7_2.Rising_Pulse_2,
           Memory_Bit_1             := "DB SENSOR CHECK".B7_2.Memory_Bit_1,
           Memory_Bit_2             := "DB SENSOR CHECK".B7_2.Memory_Bit_2,
           Word_Buffer              := "DB SENSOR CHECK".B7_2.Word_buffer,
           Word_Result              := "DB SENSOR CHECK".B7_2.Word_Result);

NETWORK
TITLE =
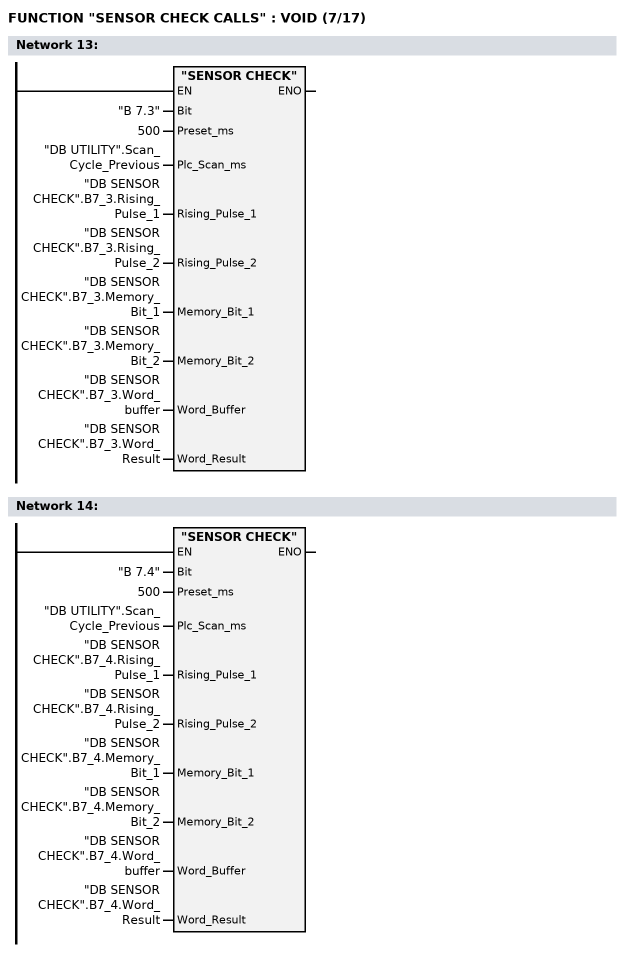

      CALL "SENSOR CHECK" (
           Bit                      := "B 7.3",
           Preset_ms                := 500,
           Plc_Scan_ms              := "DB UTILITY".Scan_Cycle_Previous,
           Rising_Pulse_1           := "DB SENSOR CHECK".B7_3.Rising_Pulse_1,
           Rising_Pulse_2           := "DB SENSOR CHECK".B7_3.Rising_Pulse_2,
           Memory_Bit_1             := "DB SENSOR CHECK".B7_3.Memory_Bit_1,
           Memory_Bit_2             := "DB SENSOR CHECK".B7_3.Memory_Bit_2,
           Word_Buffer              := "DB SENSOR CHECK".B7_3.Word_buffer,
           Word_Result              := "DB SENSOR CHECK".B7_3.Word_Result);

NETWORK
TITLE =

      CALL "SENSOR CHECK" (
           Bit                      := "B 7.4",
           Preset_ms                := 500,
           Plc_Scan_ms              := "DB UTILITY".Scan_Cycle_Previous,
           Rising_Pulse_1           := "DB SENSOR CHECK".B7_4.Rising_Pulse_1,
           Rising_Pulse_2           := "DB SENSOR CHECK".B7_4.Rising_Pulse_2,
           Memory_Bit_1             := "DB SENSOR CHECK".B7_4.Memory_Bit_1,
           Memory_Bit_2             := "DB SENSOR CHECK".B7_4.Memory_Bit_2,
           Word_Buffer              := "DB SENSOR CHECK".B7_4.Word_buffer,
           Word_Result              := "DB SENSOR CHECK".B7_4.Word_Result);

NETWORK
TITLE =
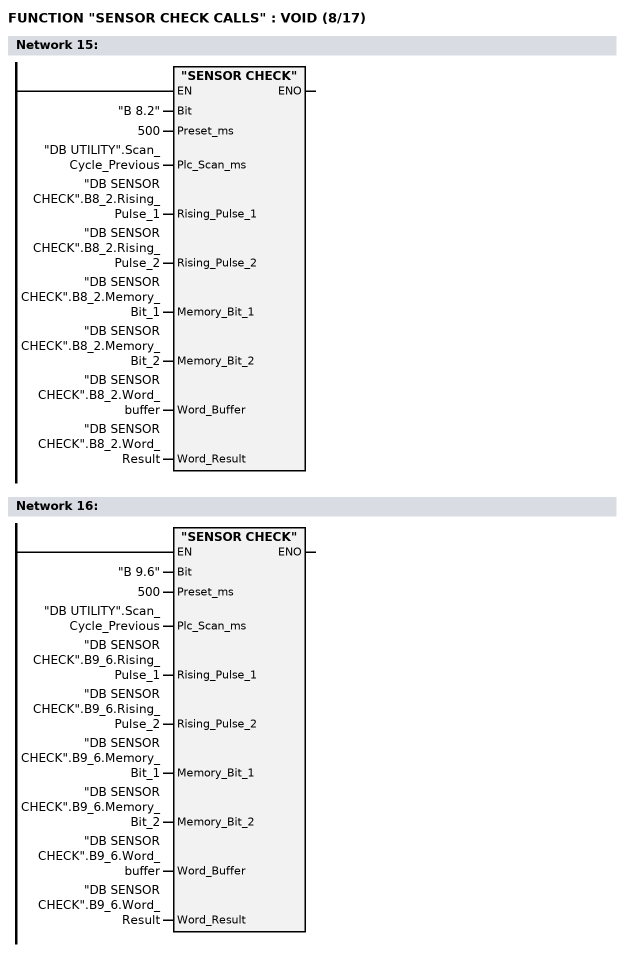

      CALL "SENSOR CHECK" (
           Bit                      := "B 8.2",
           Preset_ms                := 500,
           Plc_Scan_ms              := "DB UTILITY".Scan_Cycle_Previous,
           Rising_Pulse_1           := "DB SENSOR CHECK".B8_2.Rising_Pulse_1,
           Rising_Pulse_2           := "DB SENSOR CHECK".B8_2.Rising_Pulse_2,
           Memory_Bit_1             := "DB SENSOR CHECK".B8_2.Memory_Bit_1,
           Memory_Bit_2             := "DB SENSOR CHECK".B8_2.Memory_Bit_2,
           Word_Buffer              := "DB SENSOR CHECK".B8_2.Word_buffer,
           Word_Result              := "DB SENSOR CHECK".B8_2.Word_Result);

NETWORK
TITLE =

      CALL "SENSOR CHECK" (
           Bit                      := "B 9.6",
           Preset_ms                := 500,
           Plc_Scan_ms              := "DB UTILITY".Scan_Cycle_Previous,
           Rising_Pulse_1           := "DB SENSOR CHECK".B9_6.Rising_Pulse_1,
           Rising_Pulse_2           := "DB SENSOR CHECK".B9_6.Rising_Pulse_2,
           Memory_Bit_1             := "DB SENSOR CHECK".B9_6.Memory_Bit_1,
           Memory_Bit_2             := "DB SENSOR CHECK".B9_6.Memory_Bit_2,
           Word_Buffer              := "DB SENSOR CHECK".B9_6.Word_buffer,
           Word_Result              := "DB SENSOR CHECK".B9_6.Word_Result);

NETWORK
TITLE =
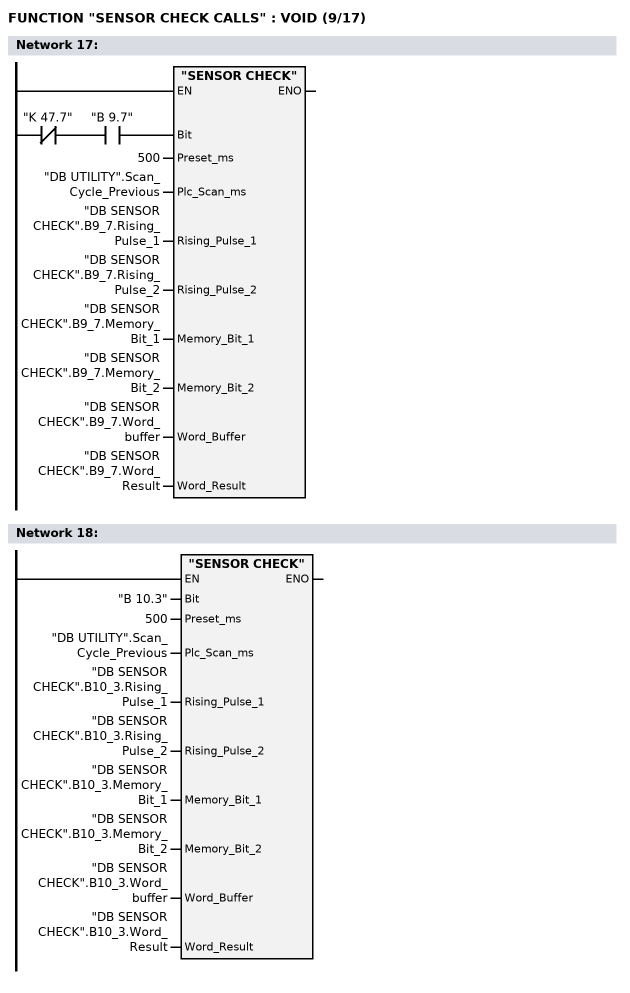

      AN    "K 47.7";
      A     "B 9.7";
      =     L      0.1;
//;
      CALL "SENSOR CHECK" (
           Bit                      := L      0.1,
           Preset_ms                := 500,
           Plc_Scan_ms              := "DB UTILITY".Scan_Cycle_Previous,
           Rising_Pulse_1           := "DB SENSOR CHECK".B9_7.Rising_Pulse_1,
           Rising_Pulse_2           := "DB SENSOR CHECK".B9_7.Rising_Pulse_2,
           Memory_Bit_1             := "DB SENSOR CHECK".B9_7.Memory_Bit_1,
           Memory_Bit_2             := "DB SENSOR CHECK".B9_7.Memory_Bit_2,
           Word_Buffer              := "DB SENSOR CHECK".B9_7.Word_buffer,
           Word_Result              := "DB SENSOR CHECK".B9_7.Word_Result);

NETWORK
TITLE =

      CALL "SENSOR CHECK" (
           Bit                      := "B 10.3",
           Preset_ms                := 500,
           Plc_Scan_ms              := "DB UTILITY".Scan_Cycle_Previous,
           Rising_Pulse_1           := "DB SENSOR CHECK".B10_3.Rising_Pulse_1,
           Rising_Pulse_2           := "DB SENSOR CHECK".B10_3.Rising_Pulse_2,
           Memory_Bit_1             := "DB SENSOR CHECK".B10_3.Memory_Bit_1,
           Memory_Bit_2             := "DB SENSOR CHECK".B10_3.Memory_Bit_2,
           Word_Buffer              := "DB SENSOR CHECK".B10_3.Word_buffer,
           Word_Result              := "DB SENSOR CHECK".B10_3.Word_Result);

NETWORK
TITLE =
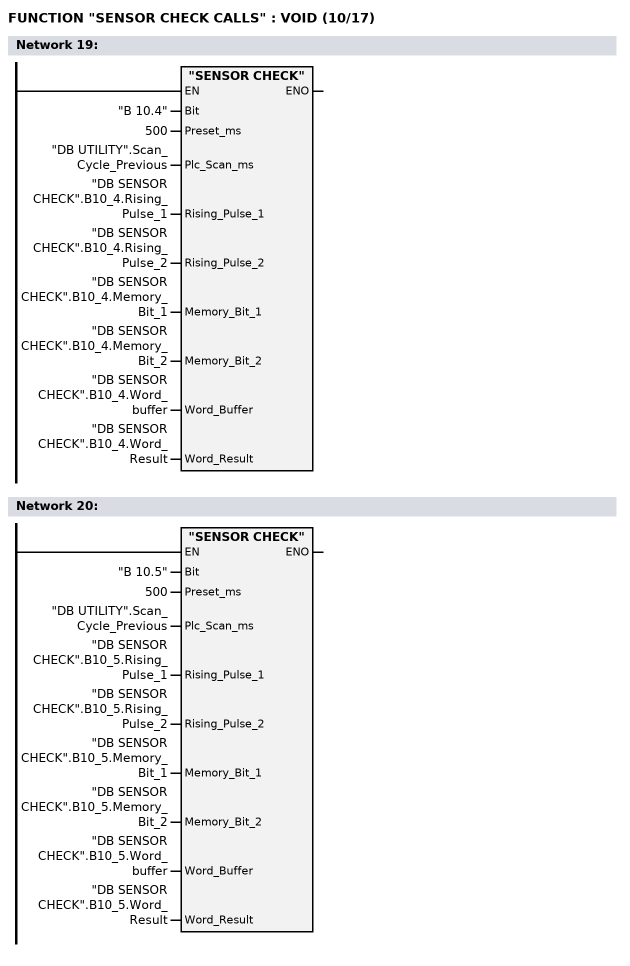

      CALL "SENSOR CHECK" (
           Bit                      := "B 10.4",
           Preset_ms                := 500,
           Plc_Scan_ms              := "DB UTILITY".Scan_Cycle_Previous,
           Rising_Pulse_1           := "DB SENSOR CHECK".B10_4.Rising_Pulse_1,
           Rising_Pulse_2           := "DB SENSOR CHECK".B10_4.Rising_Pulse_2,
           Memory_Bit_1             := "DB SENSOR CHECK".B10_4.Memory_Bit_1,
           Memory_Bit_2             := "DB SENSOR CHECK".B10_4.Memory_Bit_2,
           Word_Buffer              := "DB SENSOR CHECK".B10_4.Word_buffer,
           Word_Result              := "DB SENSOR CHECK".B10_4.Word_Result);

NETWORK
TITLE =

      CALL "SENSOR CHECK" (
           Bit                      := "B 10.5",
           Preset_ms                := 500,
           Plc_Scan_ms              := "DB UTILITY".Scan_Cycle_Previous,
           Rising_Pulse_1           := "DB SENSOR CHECK".B10_5.Rising_Pulse_1,
           Rising_Pulse_2           := "DB SENSOR CHECK".B10_5.Rising_Pulse_2,
           Memory_Bit_1             := "DB SENSOR CHECK".B10_5.Memory_Bit_1,
           Memory_Bit_2             := "DB SENSOR CHECK".B10_5.Memory_Bit_2,
           Word_Buffer              := "DB SENSOR CHECK".B10_5.Word_buffer,
           Word_Result              := "DB SENSOR CHECK".B10_5.Word_Result);

NETWORK
TITLE =
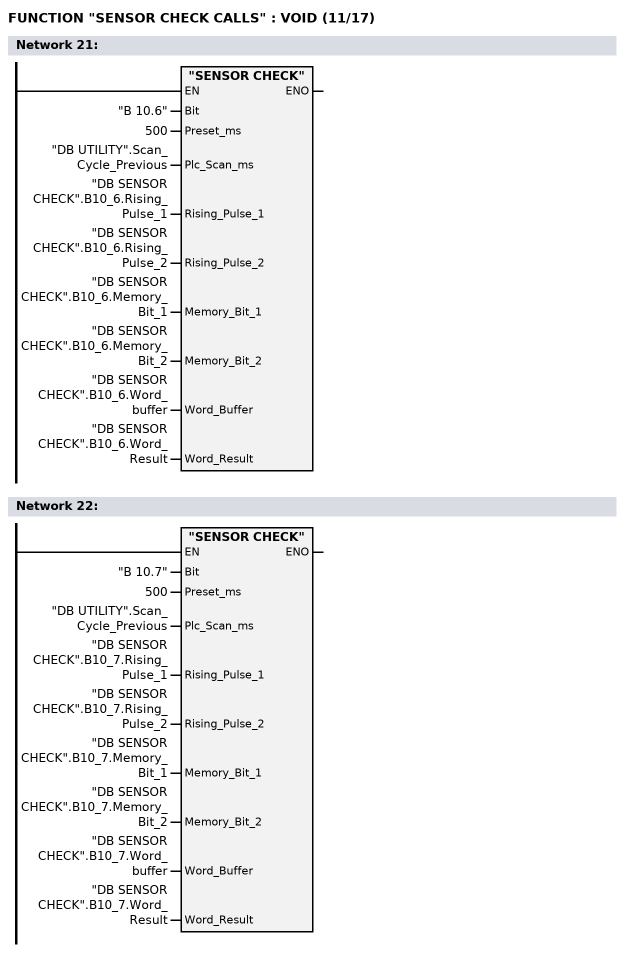

      CALL "SENSOR CHECK" (
           Bit                      := "B 10.6",
           Preset_ms                := 500,
           Plc_Scan_ms              := "DB UTILITY".Scan_Cycle_Previous,
           Rising_Pulse_1           := "DB SENSOR CHECK".B10_6.Rising_Pulse_1,
           Rising_Pulse_2           := "DB SENSOR CHECK".B10_6.Rising_Pulse_2,
           Memory_Bit_1             := "DB SENSOR CHECK".B10_6.Memory_Bit_1,
           Memory_Bit_2             := "DB SENSOR CHECK".B10_6.Memory_Bit_2,
           Word_Buffer              := "DB SENSOR CHECK".B10_6.Word_buffer,
           Word_Result              := "DB SENSOR CHECK".B10_6.Word_Result);

NETWORK
TITLE =

      CALL "SENSOR CHECK" (
           Bit                      := "B 10.7",
           Preset_ms                := 500,
           Plc_Scan_ms              := "DB UTILITY".Scan_Cycle_Previous,
           Rising_Pulse_1           := "DB SENSOR CHECK".B10_7.Rising_Pulse_1,
           Rising_Pulse_2           := "DB SENSOR CHECK".B10_7.Rising_Pulse_2,
           Memory_Bit_1             := "DB SENSOR CHECK".B10_7.Memory_Bit_1,
           Memory_Bit_2             := "DB SENSOR CHECK".B10_7.Memory_Bit_2,
           Word_Buffer              := "DB SENSOR CHECK".B10_7.Word_buffer,
           Word_Result              := "DB SENSOR CHECK".B10_7.Word_Result);

NETWORK
TITLE =
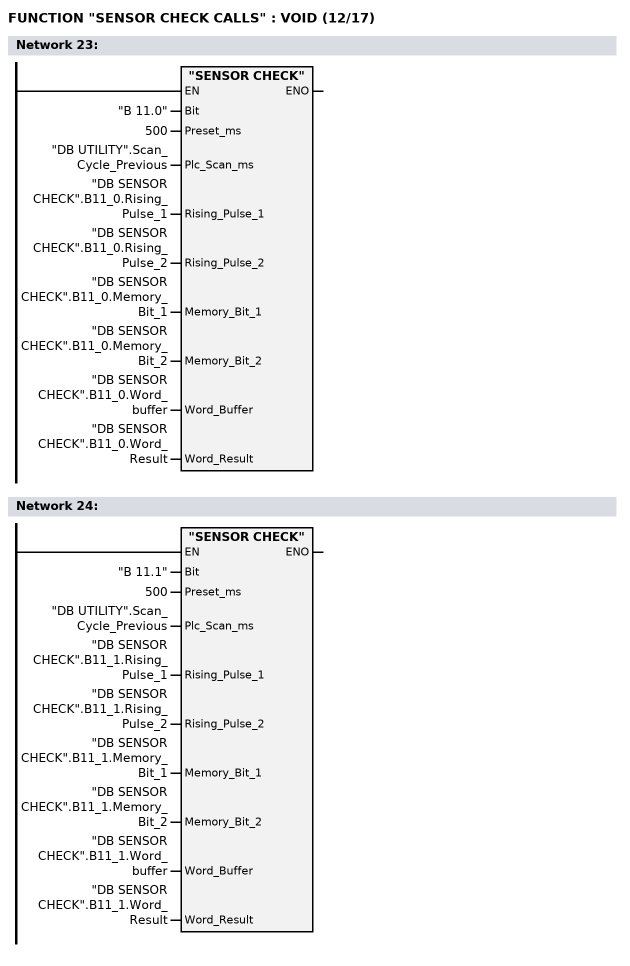

      CALL "SENSOR CHECK" (
           Bit                      := "B 11.0",
           Preset_ms                := 500,
           Plc_Scan_ms              := "DB UTILITY".Scan_Cycle_Previous,
           Rising_Pulse_1           := "DB SENSOR CHECK".B11_0.Rising_Pulse_1,
           Rising_Pulse_2           := "DB SENSOR CHECK".B11_0.Rising_Pulse_2,
           Memory_Bit_1             := "DB SENSOR CHECK".B11_0.Memory_Bit_1,
           Memory_Bit_2             := "DB SENSOR CHECK".B11_0.Memory_Bit_2,
           Word_Buffer              := "DB SENSOR CHECK".B11_0.Word_buffer,
           Word_Result              := "DB SENSOR CHECK".B11_0.Word_Result);

NETWORK
TITLE =

      CALL "SENSOR CHECK" (
           Bit                      := "B 11.1",
           Preset_ms                := 500,
           Plc_Scan_ms              := "DB UTILITY".Scan_Cycle_Previous,
           Rising_Pulse_1           := "DB SENSOR CHECK".B11_1.Rising_Pulse_1,
           Rising_Pulse_2           := "DB SENSOR CHECK".B11_1.Rising_Pulse_2,
           Memory_Bit_1             := "DB SENSOR CHECK".B11_1.Memory_Bit_1,
           Memory_Bit_2             := "DB SENSOR CHECK".B11_1.Memory_Bit_2,
           Word_Buffer              := "DB SENSOR CHECK".B11_1.Word_buffer,
           Word_Result              := "DB SENSOR CHECK".B11_1.Word_Result);

NETWORK
TITLE =
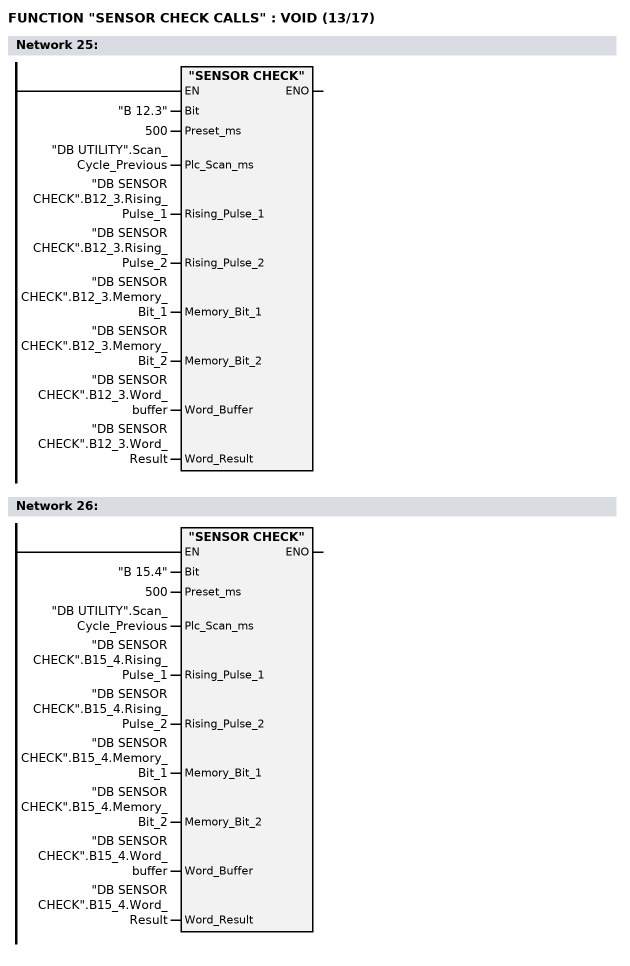

      CALL "SENSOR CHECK" (
           Bit                      := "B 12.3",
           Preset_ms                := 500,
           Plc_Scan_ms              := "DB UTILITY".Scan_Cycle_Previous,
           Rising_Pulse_1           := "DB SENSOR CHECK".B12_3.Rising_Pulse_1,
           Rising_Pulse_2           := "DB SENSOR CHECK".B12_3.Rising_Pulse_2,
           Memory_Bit_1             := "DB SENSOR CHECK".B12_3.Memory_Bit_1,
           Memory_Bit_2             := "DB SENSOR CHECK".B12_3.Memory_Bit_2,
           Word_Buffer              := "DB SENSOR CHECK".B12_3.Word_buffer,
           Word_Result              := "DB SENSOR CHECK".B12_3.Word_Result);

NETWORK
TITLE =

      CALL "SENSOR CHECK" (
           Bit                      := "B 15.4",
           Preset_ms                := 500,
           Plc_Scan_ms              := "DB UTILITY".Scan_Cycle_Previous,
           Rising_Pulse_1           := "DB SENSOR CHECK".B15_4.Rising_Pulse_1,
           Rising_Pulse_2           := "DB SENSOR CHECK".B15_4.Rising_Pulse_2,
           Memory_Bit_1             := "DB SENSOR CHECK".B15_4.Memory_Bit_1,
           Memory_Bit_2             := "DB SENSOR CHECK".B15_4.Memory_Bit_2,
           Word_Buffer              := "DB SENSOR CHECK".B15_4.Word_buffer,
           Word_Result              := "DB SENSOR CHECK".B15_4.Word_Result);

NETWORK
TITLE =
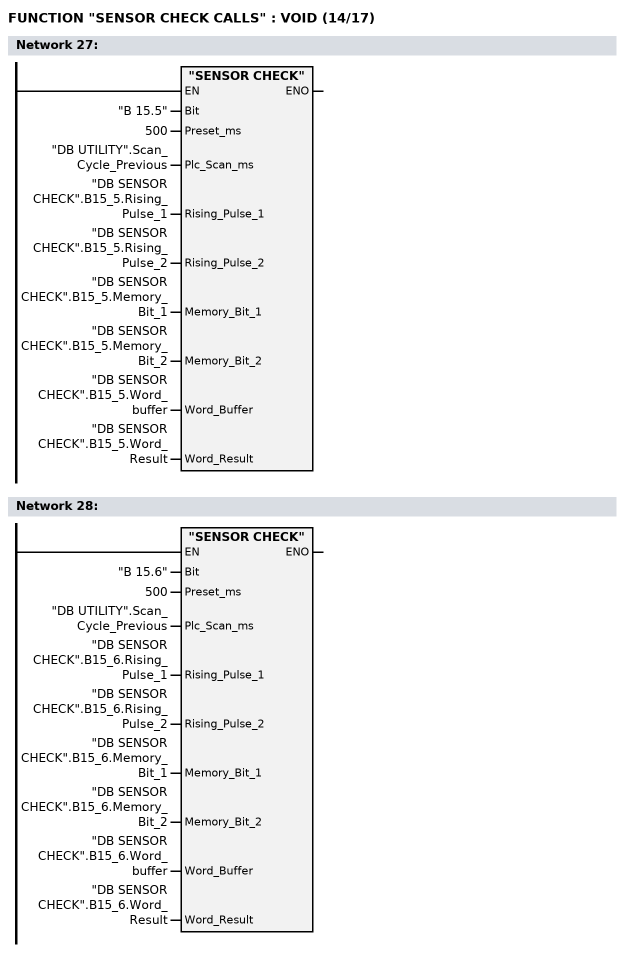

      CALL "SENSOR CHECK" (
           Bit                      := "B 15.5",
           Preset_ms                := 500,
           Plc_Scan_ms              := "DB UTILITY".Scan_Cycle_Previous,
           Rising_Pulse_1           := "DB SENSOR CHECK".B15_5.Rising_Pulse_1,
           Rising_Pulse_2           := "DB SENSOR CHECK".B15_5.Rising_Pulse_2,
           Memory_Bit_1             := "DB SENSOR CHECK".B15_5.Memory_Bit_1,
           Memory_Bit_2             := "DB SENSOR CHECK".B15_5.Memory_Bit_2,
           Word_Buffer              := "DB SENSOR CHECK".B15_5.Word_buffer,
           Word_Result              := "DB SENSOR CHECK".B15_5.Word_Result);

NETWORK
TITLE =

      CALL "SENSOR CHECK" (
           Bit                      := "B 15.6",
           Preset_ms                := 500,
           Plc_Scan_ms              := "DB UTILITY".Scan_Cycle_Previous,
           Rising_Pulse_1           := "DB SENSOR CHECK".B15_6.Rising_Pulse_1,
           Rising_Pulse_2           := "DB SENSOR CHECK".B15_6.Rising_Pulse_2,
           Memory_Bit_1             := "DB SENSOR CHECK".B15_6.Memory_Bit_1,
           Memory_Bit_2             := "DB SENSOR CHECK".B15_6.Memory_Bit_2,
           Word_Buffer              := "DB SENSOR CHECK".B15_6.Word_buffer,
           Word_Result              := "DB SENSOR CHECK".B15_6.Word_Result);

NETWORK
TITLE =
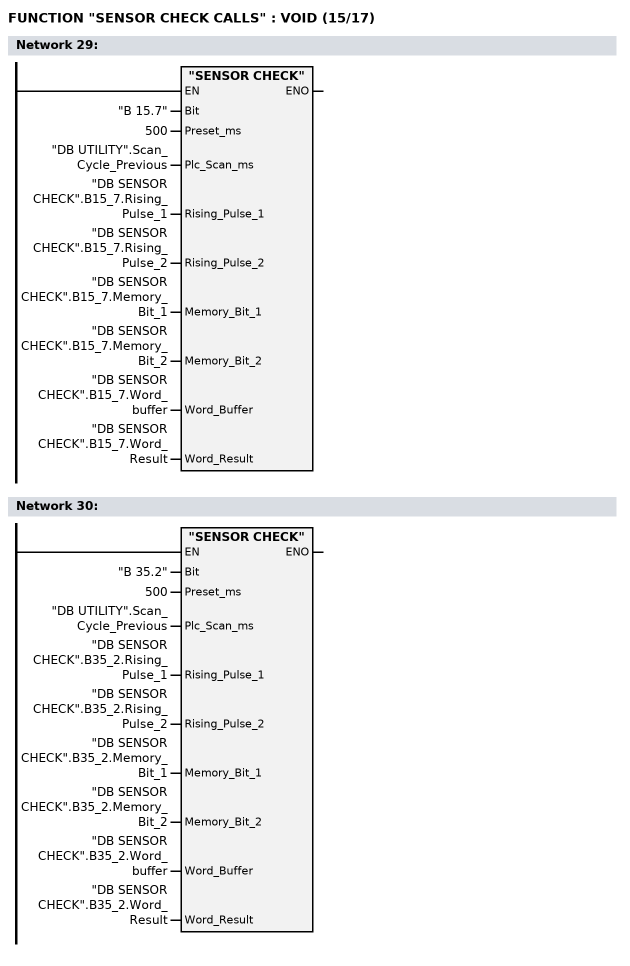

      CALL "SENSOR CHECK" (
           Bit                      := "B 15.7",
           Preset_ms                := 500,
           Plc_Scan_ms              := "DB UTILITY".Scan_Cycle_Previous,
           Rising_Pulse_1           := "DB SENSOR CHECK".B15_7.Rising_Pulse_1,
           Rising_Pulse_2           := "DB SENSOR CHECK".B15_7.Rising_Pulse_2,
           Memory_Bit_1             := "DB SENSOR CHECK".B15_7.Memory_Bit_1,
           Memory_Bit_2             := "DB SENSOR CHECK".B15_7.Memory_Bit_2,
           Word_Buffer              := "DB SENSOR CHECK".B15_7.Word_buffer,
           Word_Result              := "DB SENSOR CHECK".B15_7.Word_Result);

NETWORK
TITLE =

      CALL "SENSOR CHECK" (
           Bit                      := "B 35.2",
           Preset_ms                := 500,
           Plc_Scan_ms              := "DB UTILITY".Scan_Cycle_Previous,
           Rising_Pulse_1           := "DB SENSOR CHECK".B35_2.Rising_Pulse_1,
           Rising_Pulse_2           := "DB SENSOR CHECK".B35_2.Rising_Pulse_2,
           Memory_Bit_1             := "DB SENSOR CHECK".B35_2.Memory_Bit_1,
           Memory_Bit_2             := "DB SENSOR CHECK".B35_2.Memory_Bit_2,
           Word_Buffer              := "DB SENSOR CHECK".B35_2.Word_buffer,
           Word_Result              := "DB SENSOR CHECK".B35_2.Word_Result);

NETWORK
TITLE =
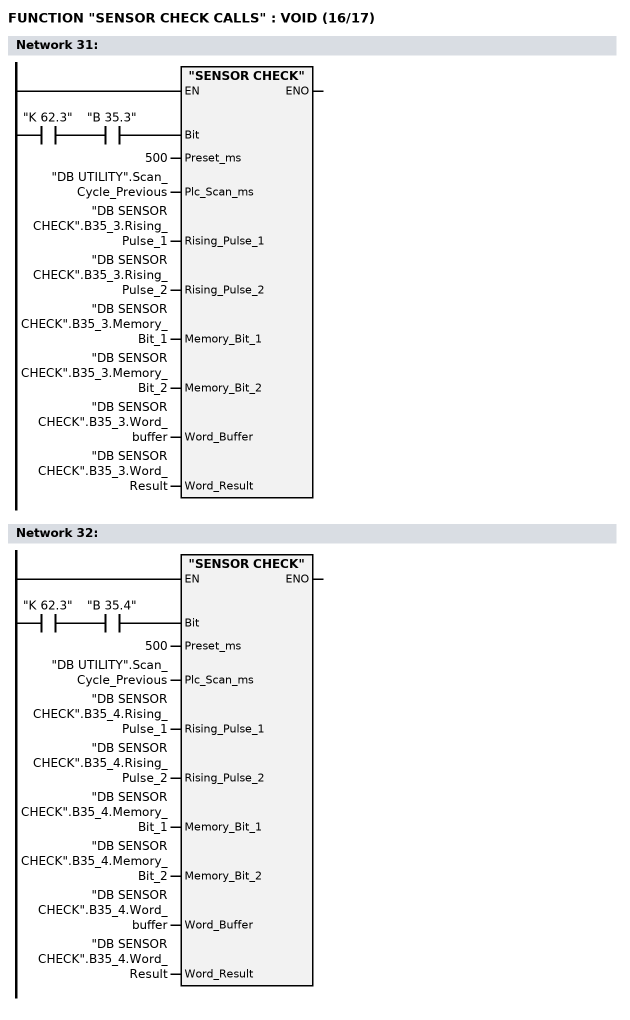

      A     "K 62.3";
      A     "B 35.3";
      =     L      0.2;

      CALL "SENSOR CHECK" (
           Bit                      := L      0.2,
           Preset_ms                := 500,
           Plc_Scan_ms              := "DB UTILITY".Scan_Cycle_Previous,
           Rising_Pulse_1           := "DB SENSOR CHECK".B35_3.Rising_Pulse_1,
           Rising_Pulse_2           := "DB SENSOR CHECK".B35_3.Rising_Pulse_2,
           Memory_Bit_1             := "DB SENSOR CHECK".B35_3.Memory_Bit_1,
           Memory_Bit_2             := "DB SENSOR CHECK".B35_3.Memory_Bit_2,
           Word_Buffer              := "DB SENSOR CHECK".B35_3.Word_buffer,
           Word_Result              := "DB SENSOR CHECK".B35_3.Word_Result);

NETWORK
TITLE =

      A     "K 62.3";
      A     "B 35.4";
      =     L      0.3;
//;
      CALL "SENSOR CHECK" (
           Bit                      := L      0.3,
           Preset_ms                := 500,
           Plc_Scan_ms              := "DB UTILITY".Scan_Cycle_Previous,
           Rising_Pulse_1           := "DB SENSOR CHECK".B35_4.Rising_Pulse_1,
           Rising_Pulse_2           := "DB SENSOR CHECK".B35_4.Rising_Pulse_2,
           Memory_Bit_1             := "DB SENSOR CHECK".B35_4.Memory_Bit_1,
           Memory_Bit_2             := "DB SENSOR CHECK".B35_4.Memory_Bit_2,
           Word_Buffer              := "DB SENSOR CHECK".B35_4.Word_buffer,
           Word_Result              := "DB SENSOR CHECK".B35_4.Word_Result);

NETWORK
TITLE =
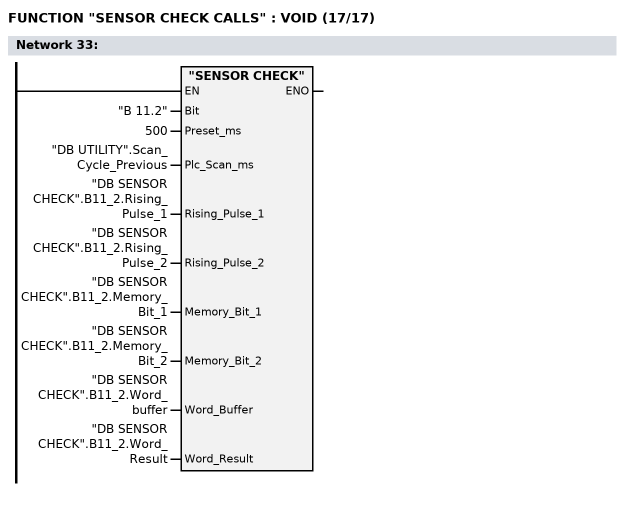

      CALL "SENSOR CHECK" (
           Bit                      := "B 11.2",
           Preset_ms                := 500,
           Plc_Scan_ms              := "DB UTILITY".Scan_Cycle_Previous,
           Rising_Pulse_1           := "DB SENSOR CHECK".B11_2.Rising_Pulse_1,
           Rising_Pulse_2           := "DB SENSOR CHECK".B11_2.Rising_Pulse_2,
           Memory_Bit_1             := "DB SENSOR CHECK".B11_2.Memory_Bit_1,
           Memory_Bit_2             := "DB SENSOR CHECK".B11_2.Memory_Bit_2,
           Word_Buffer              := "DB SENSOR CHECK".B11_2.Word_buffer,
           Word_Result              := "DB SENSOR CHECK".B11_2.Word_Result);

END_FUNCTION

FUNCTION "LAUER_RE-START_PUP" : VOID
TITLE =
//Logique de remise à zéro du bit de redémarrage de la communication avec
//l'interface.
//
//Ce bit doit être remis à zéro en cas de perte de communication avec l'automate
//ou si l'interface est éteint.
VERSION : 0.1

BEGIN
NETWORK
TITLE =Lauer restart bit
//DB50.DBW25 = S and mS   “Start a 5-second watchdog timer unless reset is
//active”
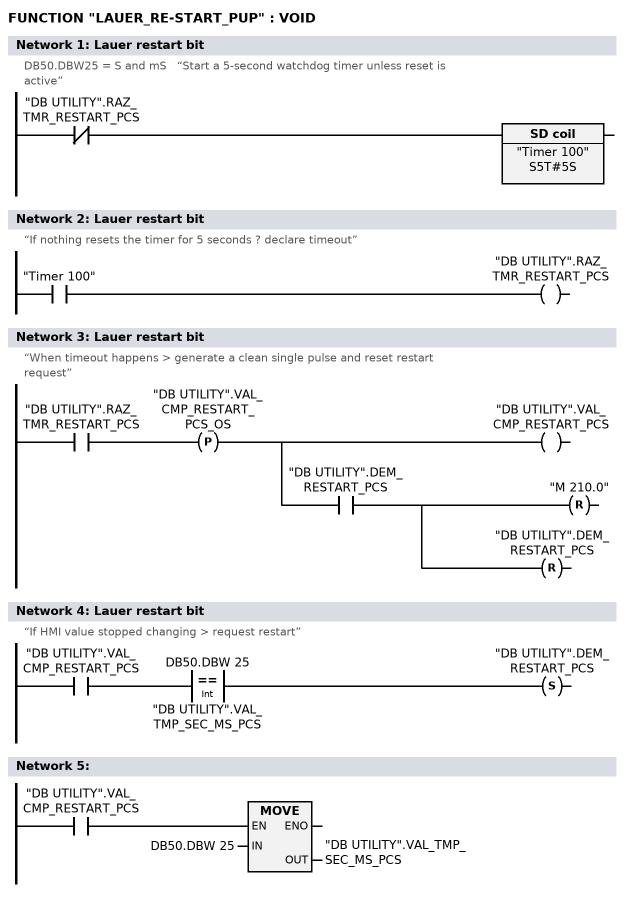
      AN    "DB UTILITY".RAZ_TMR_RESTART_PCS;
      L     S5T#5S;
      SD    "Timer 100";
      NOP   0;
      NOP   0;
      NOP   0;
      NOP   0;
NETWORK
TITLE =Lauer restart bit
//“If nothing resets the timer for 5 seconds ? declare timeout”
      A     "Timer 100";
      =     "DB UTILITY".RAZ_TMR_RESTART_PCS;
NETWORK
TITLE =Lauer restart bit
//“When timeout happens > generate a clean single pulse and reset restart
//request”
      A     "DB UTILITY".RAZ_TMR_RESTART_PCS;
      FP    "DB UTILITY".VAL_CMP_RESTART_PCS_OS;
      =     L      0.0;
      A     L      0.0;
      BLD   102;
      =     "DB UTILITY".VAL_CMP_RESTART_PCS;
      A     L      0.0;
      A     "DB UTILITY".DEM_RESTART_PCS;
      R     "M 210.0";
      R     "DB UTILITY".DEM_RESTART_PCS;
NETWORK
TITLE =Lauer restart bit
//“If HMI value stopped changing > request restart”
      A     "DB UTILITY".VAL_CMP_RESTART_PCS;
      A(    ;
      L     DB50.DBW   25;
      L     "DB UTILITY".VAL_TMP_SEC_MS_PCS;
      ==I   ;
      )     ;
      S     "DB UTILITY".DEM_RESTART_PCS;
NETWORK
TITLE =

      A     "DB UTILITY".VAL_CMP_RESTART_PCS;
      JNB   _001;
      L     DB50.DBW   25;
      T     "DB UTILITY".VAL_TMP_SEC_MS_PCS;
_001: NOP   0;
END_FUNCTION

FUNCTION "LAUER COMM ERR FC" : VOID
TITLE =
VERSION : 0.1

BEGIN
NETWORK
TITLE =
//;    Please choose your PCS and add the commands to your network
//;                      // Example PCS900/PCS 920/PCS950
//;                      // Typical presets
//;L W#16#1F00;  //(3F00 PCS950/PCS 920)
//;T DBW 72;
//;L W#16#00FF;
//;T DBW 74;
//;L W#16#0080;
//:T DBW 76;
//;                      // Example PCS009/PCS090/PCS095
//;                      // Typical presets
//;     L W#16#0FC8;
//;     T DBW 26;
//;     L W#16#0080;
//;     T DBW 28;
      L     W#16#0;
      T     DBW    8;
      T     DBW   10;
      T     DBW   12;
      T     DBW   14;
      T     DBW   46;
END_FUNCTION

FUNCTION "LAUER RESTART FC" : VOID
TITLE =
NAME : COFF
VERSION : 0.0

BEGIN
NETWORK
TITLE =
//;                     // Presets emergancy case
//;// Clear all keys
      L     W#16#0;
      T     DBW    8;
      T     DBW   10;
      T     DBW   12;
      T     DBW   14;
      T     DBW   46;
END_FUNCTION

FUNCTION "LAUER COMM FC" : VOID
TITLE =Handling Block Profibus
//
NAME : PROFIBUS
VERSION : 0.0


VAR_INPUT
  UBDB : BLOCK_DB ;	// UBDB
  RXFA : INT ;	// RXFA
  RXLE : INT ;	// RXLE
  TXFA : INT ;	// TXFA
  TXLE : INT ;	// TXLE
  RSET : BOOL ;	// RSET
  TIMT : TIMER ;	// TIMT
  TIMZ : S5TIME ;	// TIMZ
  COFF : BLOCK_FC ;	// COFF
  INIT : BLOCK_FC ;	// INIT
END_VAR
VAR_OUTPUT
  RFLM : BOOL ;	// RFLM
  EROR : BOOL ;	// EROR
END_VAR
VAR_TEMP
  conv_akku1 : DWORD ;
  conv_akku2 : DWORD ;
  conv_stw : WORD ;
END_VAR
BEGIN
NETWORK
TITLE =

      OPN   #UBDB; //  --------------------------
      AN    #RFLM; //  First action in FB?
      JC    OK;
      A     #TIMT; //  Timeout and no restart?
      AN    #RSET;
      JC    ERR;
      A     #TIMT;
      AN    #EROR;
      JC    ERR;
      JU    OK;

ERR:  A     #EROR;
      JC    ERR1;
      UC    #COFF; //  Call COFF once.
      OPN   #UBDB;

ERR1: A     #TIMT; //  If timeout set error-flag.
      S     #EROR;
      BEU   ;

OK:   A     #RFLM; //  First action?
      JC    CONT;
      UC    #INIT; //  Call INIT once.
      OPN   #UBDB;
      L     W#16#0; //  Init ----------------------
      T     DBW    0;
      T     DBW    2;
      T     DBW    4;
      T     DBW    6;
      AN    #RFLM;
      S     #RFLM; //  Set reset-ready-flag
//;
      AN    #RFLM; //  Trigger timer
      L     #TIMZ;
      SD    #TIMT;
//;
      A     #RFLM;
      L     #TIMZ;
      SD    #TIMT;

CONT: L     #RXFA;
      T     "MW 244"; //  ----------------------------
      +     1; //  Adress Handle1 E-Box
      T     "MW 252";
      L     #RXLE; //  Adress of first instruction
      +     -2;
      T     "MW 250"; //  Lenght E-Box Userdatas
//;
      L     #TXFA;
      T     "MW 242";
      +     1; //  Adress Handle1 A-Box
      T     "MW 248";
      L     #TXLE; //  Adress of first senddata
      +     -2;
      T     "MW 246"; //  Lenght A-Box-Userdatas
//;
      L     "MW 244"; //  Handle2 != Handle1? ---------
      L     #RXLE;
      +I    ;
      +     -1;
      T     "MW 238"; //  Adress Handle2
      T     #conv_akku1;
//;
      L     STW;
      T     #conv_stw;
//;
      L     "MB 239";
      SLW   3;
      LAR1  ;
      L     #conv_stw;
      T     STW;
//;
      L     #conv_akku1;
      L     IB [AR1,P#0.0];
      T     "MW 238"; //  Handle2
      T     #conv_akku1; //  Adress Handle1
//;
      L     STW;
      T     #conv_stw;
//;
      L     "MB 245";
      SLW   3;
      LAR1  ;
      L     #conv_stw;
      T     STW;
//;
      L     #conv_akku1;
      L     IB [AR1,P#0.0];
      L     "MW 238";
      <>I   ;
      BEC   ; //  Handle1 != Handle2 -> EXIT
//;
      T     #conv_akku1; //  Handle1 != HandleAlt? -------

      L     STW;
      T     #conv_stw;
//;
      L     "MB 245";
      SLW   3;
      LAR1  ;
      L     #conv_stw;
      T     STW;
//;
      L     #conv_akku1;
      L     IB [AR1,P#0.0];
      L     DBW    0; //  HandleAlt in UBDB (0)
      ==I   ;
      BEC   ;
//;
      AN    #RFLM; //  Start timeout-timer
      L     #TIMZ;
      SD    #TIMT;
//;
      A     #RFLM;
      L     #TIMZ;
      SD    #TIMT;
//;
      T     #conv_akku1; //  First action requiered?
      L     STW;
      T     #conv_stw;
      L     "MB 245";
      SLW   3;
      LAR1  ;
      L     #conv_stw;
      T     STW;
//;
      L     #conv_akku1;
      L     IB [AR1,P#0.0];
      L     W#16#80; //  Handle == 0x80?
      <>I   ;
      JC    SLP1;
      A     #RSET; // Clear Restart-Flag.
      R     #RSET;

END:  NOP   0;

      T     #conv_akku1; // Get Handle1(E) from RX-Box.

      L     STW;
      T     #conv_stw;
//;
      L     "MB 245";
      SLW   3;
      LAR1  ;
      L     #conv_stw;
      T     STW;
//;
      L     #conv_akku1;
      L     IB [AR1,P#0.0];
      T     DBW    0; // Save to HandleAlt.
      INVI  ; // Invert.
      T     "MW 236"; // Temporary saved.
      L     "MW 236";
      T     #conv_akku1; // Take inverted Handle1(E) to
      TAK   ;
      T     #conv_akku2;
      L     STW;
      T     #conv_stw;
//;
      L     "MB 243";
      SLW   3;
      LAR1  ;
      L     #conv_stw;
      T     STW;
//;
      L     #conv_akku2;
      L     #conv_akku1;
      T     QB [AR1,P#0.0]; // Handle1(A).
//;
      L     "MW 242";
      L     #TXLE;
      +I    ;
      +     -1;
      T     "MW 238"; // Take inverted Handle1(E) to
      L     "MW 236";
      T     #conv_akku1;
      TAK   ;
      T     #conv_akku2;
      L     STW;
      T     #conv_stw;
//;
      L     "MB 239";
      SLW   3;
      LAR1  ;
      L     #conv_stw;
      T     STW;
//;
      L     #conv_akku2;
      L     #conv_akku1;
      T     QB [AR1,P#0.0];
//;
      AN    #TIMT; // Clear Error-Mark.
      R     #EROR;
      BEU   ; // see you later...

SLP1: L     #RXFA; // Reached Rx-Box-End?
      L     #RXLE;
      +I    ;
      +     -1;
      L     "MW 252";
      ==I   ;
      JC    END;

      T     #conv_akku1; //  Start/Continue--------------

      L     STW;
      T     #conv_stw;
//;
      L     "MB 253";
      SLW   3;
      LAR1  ;
      L     #conv_stw;
      T     STW;
//;
      L     #conv_akku1;
      L     IW [AR1,P#0.0];
      L     W#16#0; //  Is anything usable?
      ==I   ;
      JC    END;

      T     #conv_akku1; //  Get first ABW.

      L     STW;
      T     #conv_stw;
//;
      L     "MB 253";
      SLW   3;
      LAR1  ;
      L     #conv_stw;
      T     STW;
//;
      L     #conv_akku1;
      L     IB [AR1,P#0.0];
      T     "MW 240"; //  Adress(UBDB) in ABW.
      L     "MW 252";
      +     1; //  Increment RX-Pointer.
      T     "MW 252";
      T     #conv_akku1;
      L     STW;
      T     #conv_stw;
      L     "MB 253";
      SLW   3;
      LAR1  ;
      L     #conv_stw;
      T     STW;
//;
      L     #conv_akku1;
      L     IB [AR1,P#0.0]; //  Count of ABW: Bit3..0.
      T     "MW 238"; //  Command of ABW: Bit 7..4.
      L     "MW 252"; //  ABW pointer to next ABW
      +     1; //  or first data.
      T     "MW 252";
//;
      L     "MW 238"; //  Check for right command.
      L     W#16#F0;
      AW    ;
      T     "MW 236"; //  Temporary saved.
//;
      L     "MW 236";
      L     W#16#10;
      ==I   ;
      JC    IOK;
//;
      L     "MW 236";
      L     W#16#20;
      ==I   ;
      JC    IOK;
//;
      L     "MW 236";
      L     W#16#40;
      ==I   ;
      JC    IOK;
//;
      L     "MW 236";
      L     W#16#80;
      ==I   ;
      JC    IOK;
      BEU   ; //  Command is wrong!
//;
IOK:  L     "MW 238"; //  Command is ok.
SLP2: L     W#16#F;
      AW    ; //  Count == 0:
      JZ    SLP1; //  Next subpaket
//;
      AN    "M 239.4";
      JC    ELS1;
      OPN   #UBDB;

      T     #conv_akku1; //  Offset ABW Adress in UBDB

      L     STW;
      T     #conv_stw;
//;
      L     "MB 241";
      SLW   4;
      LAR1  ;
      L     #conv_stw;
      T     STW;
//;
      L     #conv_akku1;
      L     DBW [AR1,P#0.0];
      T     #conv_akku1; //  Pointer to TX-Box
      TAK   ;
      T     #conv_akku2;
      L     STW;
      T     #conv_stw;
//;
      L     "MB 249";
      SLW   3;
      LAR1  ;
      L     #conv_stw;
      T     STW;
//;
      L     #conv_akku2;
      L     #conv_akku1;
      T     QW [AR1,P#0.0]; //  Write to TX-Box.
      L     "MW 248";
      +     2;
      T     "MW 248";
      JU    COMM;

ELS1: NOP   0;

      T     #conv_akku1; //  Pointer to RX-Box.

      L     STW;
      T     #conv_stw;
//;
      L     "MB 253";
      SLW   3;
      LAR1  ;
      L     #conv_stw;
      T     STW;
//;
      L     #conv_akku1;
      L     IW [AR1,P#0.0];
      T     "MW 236"; //  Read Data/Mask from RX-Box.
      L     "MW 252"; //  Increment Pointer to RX-Box.
      +     2;
      T     "MW 252";
//;
      AN    "M 239.5"; //  WRITE/(AND/OR)
      JC    ELS2;
      L     "MW 236";
      OPN   #UBDB;

      T     #conv_akku1; //  Offset ABW Adress in UBDB.
      TAK   ;
      T     #conv_akku2;
      L     STW;
      T     #conv_stw;
      L     "MB 241";
      SLW   4;
      LAR1  ;
      L     #conv_stw;
      T     STW;
//;
      L     #conv_akku2;
      L     #conv_akku1;
      T     DBW [AR1,P#0.0]; //  Write to UBDB.
      JU    COMM;

ELS2: AN    "M 239.6";
      JC    ELS3;
      L     "MW 236";
      OPN   #UBDB;

      T     #conv_akku1; //  Offset ABW Adress in UBDB.
      L     STW;
      T     #conv_stw;
      L     "MB 241";
      SLW   4;
      LAR1  ;
      L     #conv_stw;
      T     STW;
//;
      L     #conv_akku1;
      L     DBW [AR1,P#0.0];
      AW    ;
      OPN   #UBDB;
      T     #conv_akku1;
      TAK   ;
      T     #conv_akku2;
      L     STW;
      T     #conv_stw;
      L     "MB 241";
      SLW   4;
      LAR1  ;
      L     #conv_stw;
      T     STW;
//;
      L     #conv_akku2;
      L     #conv_akku1;
      T     DBW [AR1,P#0.0]; //  And to UBDB
      JU    COMM;

ELS3: NOP   0;

      L     "MW 236";
      OPN   #UBDB;
      T     #conv_akku1;
      L     STW;
      T     #conv_stw;
      L     "MB 241";
      SLW   4;
      LAR1  ;
      L     #conv_stw;
      T     STW;
//;
      L     #conv_akku1;
      L     DBW [AR1,P#0.0];
      OW    ;
      OPN   #UBDB;

      T     #conv_akku1;
      TAK   ;
      T     #conv_akku2;
      L     STW;
      T     #conv_stw;
      L     "MB 241";
      SLW   4;
      LAR1  ;
      L     #conv_stw;
      T     STW;
//;
      L     #conv_akku2;
      L     #conv_akku1;
      T     DBW [AR1,P#0.0];
COMM: L     "MW 240";
      +     1;
      T     "MW 240";
      L     "MW 238"; //  Decrement counter of ABW.
      +     -1;
      T     "MW 238";
      JU    SLP2;
END_FUNCTION

FUNCTION "LAUER" : VOID
TITLE =
NAME : SCHRIANZ
VERSION : 0.0


VAR_TEMP
  TEMP0 : DWORD ;
  TEMP1 : DWORD ;
  TEMP2 : WORD ;
END_VAR
BEGIN
NETWORK
TITLE =



NETWORK
TITLE =



NETWORK
TITLE =

      OPN   "DB LAUER";

NETWORK
TITLE =

      AN    "M 150.7";
      JC    M001;
      L     2#100000000;
      T     DBW   72;
M001: NOP   0;
NETWORK
TITLE =

      ON    "M 150.7";
      JC    M002;
      L     2#1;
      T     DBW   76;
M002: NOP   0;
NETWORK
TITLE =



NETWORK
TITLE =

      O(    ;
      L     DBW  300;
      L     77;
      <I    ;
      )     ;
      O(    ;
      L     DBW  300;
      L     102;
      >I    ;
      )     ;
      JC    M003;
      JU    M004;
M003: L     77;
      T     DBW  300;
M004: NOP   0;
NETWORK
TITLE =

      L     "DB LAUER".D_150;
      L     77;
      <>I   ;
      JC    M005;
      L     "MW 15";
      T     "MW 200";
      L     "MB 17";
      T     MB   202;
M005: L     DBW  300;
      L     78;
      <>I   ;
      JC    M006;
      L     "MW 19";
      T     "MW 200";
      L     "MB 21";
      T     MB   202;
M006: L     DBW  300;
      L     79;
      <>I   ;
      JC    M007;
      L     "MW 23";
      T     "MW 200";
      L     "MB 25";
      T     MB   202;
M007: L     DBW  300;
      L     80;
      <>I   ;
      JC    M008;
      L     "MW 27";
      T     "MW 200";
      L     "MB 29";
      T     MB   202;
M008: L     DBW  300;
      L     81;
      <>I   ;
      JC    M009;
      L     "MW 31";
      T     "MW 200";
      L     "MB 33";
      T     MB   202;
M009: L     DBW  300;
      L     82;
      <>I   ;
      JC    M00a;
      L     "MW 35";
      T     "MW 200";
      L     "MB 37";
      T     MB   202;
M00a: L     DBW  300;
      L     83;
      <>I   ;
      JC    M00b;
      L     "MW 39";
      T     "MW 200";
      L     "MB 41";
      T     MB   202;
M00b: L     DBW  300;
      L     84;
      <>I   ;
      JC    M00c;
      L     "MW 43";
      T     "MW 200";
      L     "MB 45";
      T     MB   202;
M00c: L     DBW  300;
      L     85;
      <>I   ;
      JC    M00d;
      L     "MW 47";
      T     "MW 200";
      L     "MB 49";
      T     MB   202;
M00d: L     DBW  300;
      L     86;
      <>I   ;
      JC    M00e;
      L     "MW 51";
      T     "MW 200";
      L     "MB 53";
      T     MB   202;
M00e: L     DBW  300;
      L     87;
      <>I   ;
      JC    M00f;
      L     "MW 55";
      T     "MW 200";
      L     "MB 57";
      T     MB   202;
M00f: L     DBW  300;
      L     88;
      <>I   ;
      JC    M010;
      L     "MW 59";
      T     "MW 200";
      L     "MB 61";
      T     MB   202;
M010: L     DBW  300;
      L     89;
      <>I   ;
      JC    M011;
      L     "MW 63";
      T     "MW 200";
      T     "MW 200";
      L     "MB 65";
      T     MB   202;
M011: L     DBW  300;
      L     90;
      <>I   ;
      JC    M012;
      L     "MW 67";
      T     "MW 200";
      L     "MB 69";
      T     MB   202;
M012: L     DBW  300;
      L     91;
      <>I   ;
      JC    M013;
      L     "MW 71";
      T     "MW 200";
      L     "MB 73";
      T     MB   202;
M013: L     DBW  300;
      L     92;
      <>I   ;
      JC    M014;
      L     "MW 75";
      T     "MW 200";
      L     "MB 77";
      T     MB   202;
M014: L     DBW  300;
      L     93;
      <>I   ;
      JC    M015;
      L     "MW 79";
      T     "MW 200";
      L     "MB 81";
      T     MB   202;
M015: L     DBW  300;
      L     94;
      <>I   ;
      JC    M016;
      L     "MW 83";
      T     "MW 200";
      L     "MB 85";
      T     MB   202;
M016: L     DBW  300;
      L     95;
      <>I   ;
      JC    M017;
      L     "MW 87";
      T     "MW 200";
      L     "MB 89";
      T     MB   202;
M017: L     DBW  300;
      L     96;
      <>I   ;
      JC    M018;
      L     "MW 91";
      T     "MW 200";
      L     "MB 93";
      T     MB   202;
M018: L     DBW  300;
      L     97;
      <>I   ;
      JC    M019;
      L     "MW 95";
      T     "MW 200";
      L     "MB 97";
      T     MB   202;
M019: L     DBW  300;
      L     98;
      <>I   ;
      JC    M01a;
      L     "MW 99";
      T     "MW 200";
      L     "MB 101";
      T     MB   202;
M01a: L     DBW  300;
      L     99;
      <>I   ;
      JC    M01b;
      L     "MW 103";
      T     "MW 200";
      L     "MB 105";
      T     MB   202;
M01b: L     DBW  300;
      L     100;
      <>I   ;
      JC    M01c;
      L     "MW 107";
      T     "MW 200";
      L     "MB 109";
      T     MB   202;
M01c: L     DBW  300;
      L     101;
      <>I   ;
      JC    M01d;
      L     "MW 111";
      L     "MW 200";
      L     "MB 113";
      T     MB   202;
M01d: L     DBW  300;
      L     102;
      <>I   ;
      JC    M01e;
      L     "MW 115";
      T     "MW 200";
      L     "MB 117";
      T     MB   202;
M01e: NOP   0;
NETWORK
TITLE =

      L     W#16#0;
      T     MB   204;
      L     W#16#80;
      T     MB   207;
NETWORK
TITLE =

      AN    "M 203.0";
      JC    M01f;
      L     25;
      T     MB   204;
M020: L     MB   203;
      SRW   1;
      T     MB   203;
      L     MB   207;
      SRW   1;
      T     "MW 207";
      AN    "M 203.0";
      JC    M021;
      L     MB   204;
      INC   1;
      T     MB   204;
M021: AN    "M 207.0";
      JC    M020;
      JU    M022;
M01f: AN    "M 202.0";
      JC    M023;
      L     17;
      T     MB   204;
M024: L     MB   202;
      SRW   1;
      T     MB   202;
      L     MB   207;
      SRW   1;
      T     MB   207;
      AN    "M 202.0";
      JC    M025;
      L     MB   204;
      INC   1;
      T     MB   204;
M025: AN    "M 207.0";
      JC    M024;
      JU    M022;
M023: AN    "M 201.0";
      JC    M026;
      L     9;
      T     MB   204;
M027: L     "MB 201";
      SRW   1;
      T     "MB 201";
      L     MB   207;
      SRW   1;
      T     MB   207;
      AN    "M 201.0";
      JC    M028;
      L     MB   204;
      INC   1;
      T     MB   204;
M028: AN    "M 207.0";
      JC    M027;
      JU    M022;
M026: AN    "M 200.0";
      JC    M022;
      L     1;
      T     MB   204;
M029: L     "MB 200";
      SRW   1;
      T     "MB 200";
      L     MB   207;
      SRW   1;
      T     MB   207;
      AN    "M 200.0";
      JC    M02a;
      L     MB   204;
      INC   1;
      T     MB   204;
M02a: AN    "M 207.0";
      JC    M029;
M022: NOP   0;
NETWORK
TITLE =



NETWORK
TITLE =

      OPN   "DB LAUER";
      L     MB   204;
      T     #TEMP0;
      TAK   ;
      T     #TEMP1;
      L     STW;
      T     #TEMP2;
      L     DBB  301;
      SLW   4;
      LAR1  ;
      L     #TEMP2;
      T     STW;
      L     #TEMP1;
      L     #TEMP0;
      T     DBW [AR1,P#0.0];
NETWORK
TITLE =



NETWORK
TITLE =

      L     "DB LAUER".D_150;
      INC   1;
      T     DBW  300;
NETWORK
TITLE =



NETWORK
TITLE =



END_FUNCTION

FUNCTION "CONTROL" : VOID
TITLE =Controls
VERSION : 0.0

BEGIN
NETWORK
TITLE =Qty Accumulation Conveyor
//  A     "M 0.3"
//      A     "M 92.0"
//      AN    "M 14.4"
//      CU    "COUNTER 4"
////;
//      A     "M 0.3"
//      A     "B 6.4"
//      CD    "COUNTER 4"
////;
//      A     "M 161.0"
//      A     "M 161.1"
//      A(
//      ON    "S 2.1"
//      O     "S 2.2"
//      )
//      R     "COUNTER 4"
//


NETWORK
TITLE =Qty Accumulation Conveyor
//      A     "M 0.3"
//      AN    "B 6.7"
//      CU    "COUNTER 5"
//      A     "M 0.3"
//      AN    "B 7.2"
//      CD    "COUNTER 5"
//      A     "M 161.0"
//      A     "M 161.1"
//      A(
//      ON    "S 2.1"
//      O     "S 2.2"
//      )
//      R     "COUNTER 5"
//


NETWORK
TITLE =Qty Flipper to Pusher
//      A     "M 0.3"
//      AN    "B 7.4"
//      CU    "COUNTER 6"
//      A     "M 0.3"
//      AN    "B 10.4"
//      CD    "COUNTER 6"
//      A     "M 161.0"
//      A     "M 161.1"
//      A(
//      ON    "S 2.1"
//      O     "S 2.2"
//      )
//      R     "COUNTER 6"
//


NETWORK
TITLE =Qty Pivot / Collator Conveyor
//      A     "M 0.3"
//      AN    "B 10.4"
//      CU    "COUNTER 7"
//      A     "M 0.3"
//      AN    "B 10.5"
//      CD    "COUNTER 7"
//      A     "M 161.0"
//      A     "M 161.1"
//      A(
//      ON    "S 2.1"
//      O     "S 2.2"
//      )
//      R     "COUNTER 7"
//


NETWORK
TITLE =Qty Bottom Accumulator
//      A     "M 0.3"
//      A     "B 10.6"
//      A     "P 15.1"
//      CU    "COUNTER 8"
//      A     "M 0.3"
//      AN    "B 11.2"
//      CD    "COUNTER 8"
//      A     "M 161.0"
//      A     "M 161.1"
//      A(
//      ON    "S 2.1"
//      O     "S 2.2"
//      )
//      R     "COUNTER 8"
//


NETWORK
TITLE =Qty Top Accumulator
//      A     "M 0.3"
//      A     "B 10.6"
//      A     "P 15.0"
//      CU    "COUNTER 9"
//      A     "M 0.3"
//      AN    "B 15.6"
//      CD    "COUNTER 9"
//      A     "M 161.1"
//      A     "M 161.1"
//      A(
//      ON    "S 2.1"
//      O     "S 2.2"
//      )
//      R     "COUNTER 9"
//


NETWORK
TITLE =Start Signal
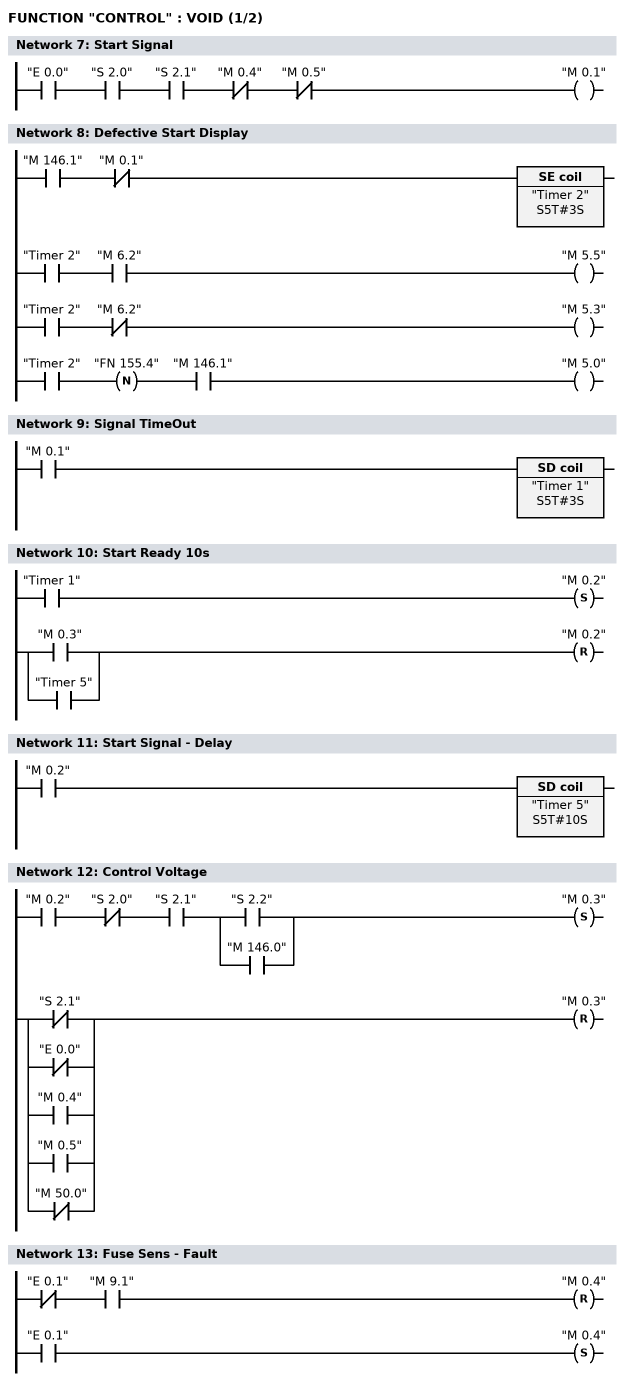

      A     "E 0.0";
      A(    ;
      O     "S 2.0";
//   O     "M 146.1"
      )     ;
      A     "S 2.1";
//      A     "M 146.2"
      AN    "M 0.4";
      AN    "M 0.5";
      =     "M 0.1";
NETWORK
TITLE =Defective Start Display

      A     "M 146.1";
      AN    "M 0.1";
      L     S5T#3S;
      SE    "Timer 2";
//;
      A     "Timer 2";
      A     "M 6.2";
      =     "M 5.5";
//;
      A     "Timer 2";
      AN    "M 6.2";
      =     "M 5.3";
//;
      A     "Timer 2";
      FN    "FN 155.4";
      A     "M 146.1";
      =     "M 5.0";
NETWORK
TITLE =Signal TimeOut

      A     "M 0.1";
      L     S5T#3S;
      SD    "Timer 1";
NETWORK
TITLE =Start Ready 10s

      A     "Timer 1";
      S     "M 0.2";
//;
      A(    ;
      O     "M 0.3";
      O     "Timer 5";
      )     ;
      R     "M 0.2";
NETWORK
TITLE =Start Signal - Delay

      A     "M 0.2";
      L     S5T#10S;
      SD    "Timer 5";
NETWORK
TITLE =Control Voltage

      A     "M 0.2";
      AN    "S 2.0";
      A     "S 2.1";
//    A    "M 146.2"
      A(    ;
      O     "S 2.2";
      O     "M 146.0";
      )     ;
      S     "M 0.3";
//;
      A(    ;
      ON    "S 2.1";
//    ON    "M 146.2"
      ON    "E 0.0";
      O     "M 0.4";
      O     "M 0.5";
      ON    "M 50.0";
      )     ;
      R     "M 0.3";
NETWORK
TITLE =Fuse Sens - Fault

      AN    "E 0.1";
      A     "M 9.1";
      R     "M 0.4";
//;
      A     "E 0.1";
      S     "M 0.4";
NETWORK
TITLE =Motor Protect - Fault
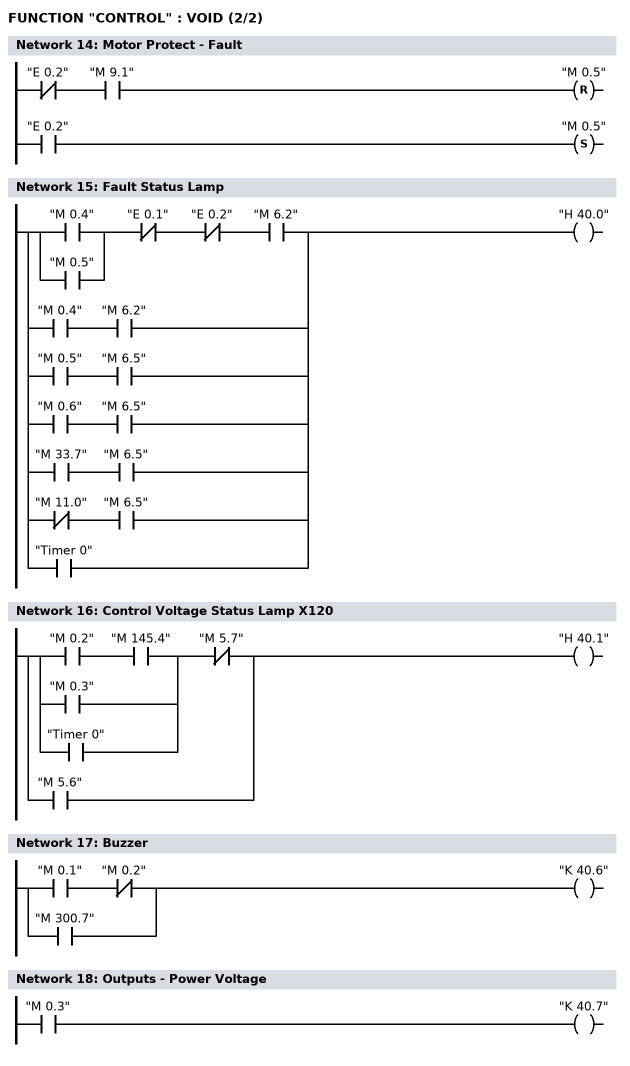

      AN    "E 0.2";
      A     "M 9.1";
      R     "M 0.5";
//;
      A     "E 0.2";
      S     "M 0.5";
NETWORK
TITLE =Fault Status Lamp

      A(    ;
      O     "M 0.4";
      O     "M 0.5";
      )     ;
      AN    "E 0.1";
      AN    "E 0.2";
      A     "M 6.2";
      O     ;
      A     "M 0.4";
      A     "M 6.2";
      O     ;
      A     "M 0.5";
      A     "M 6.5";
      O     ;
      A     "M 0.6";
      A     "M 6.5";
      O     ;
      A     "M 33.7";
      A     "M 6.5";
      O     ;
      AN    "M 11.0";
      A     "M 6.5";
      O     "Timer 0";
      =     "H 40.0";
NETWORK
TITLE =Control Voltage Status Lamp X120

      A     "M 0.2";
      A     "M 145.4";
      O     "M 0.3";
      O     "Timer 0";
      AN    "M 5.7";
      O     "M 5.6";
      =     "H 40.1";
NETWORK
TITLE =Buzzer

      A     "M 0.1";
      AN    "M 0.2";
      O     "M 300.7";
      =     "K 40.6";
NETWORK
TITLE =Outputs - Power Voltage

      A     "M 0.3";
      =     "K 40.7";
END_FUNCTION

FUNCTION "GENERAL FAULTS" : VOID
TITLE =General Faults
VERSION : 0.0


VAR_TEMP
  INIT_DELAY : BOOL ;
  CHECK_PULSE : BOOL ;
  ELEVATOR_U42_0 : BOOL ;	//CO ELEVATOR VFD U42.0 - READY    POS.2
  FAULT_TRIGGERED : BOOL ;
  FAULT_REGISTER_1 : BOOL ;
  FAULT_REGISTER_2 : BOOL ;
  FAULT_REGISTER_3 : BOOL ;
  FAULT_REGISTER_4 : BOOL ;
  FAULT_REGISTER_5 : BOOL ;
END_VAR
BEGIN
NETWORK
TITLE =Trigger Pulse
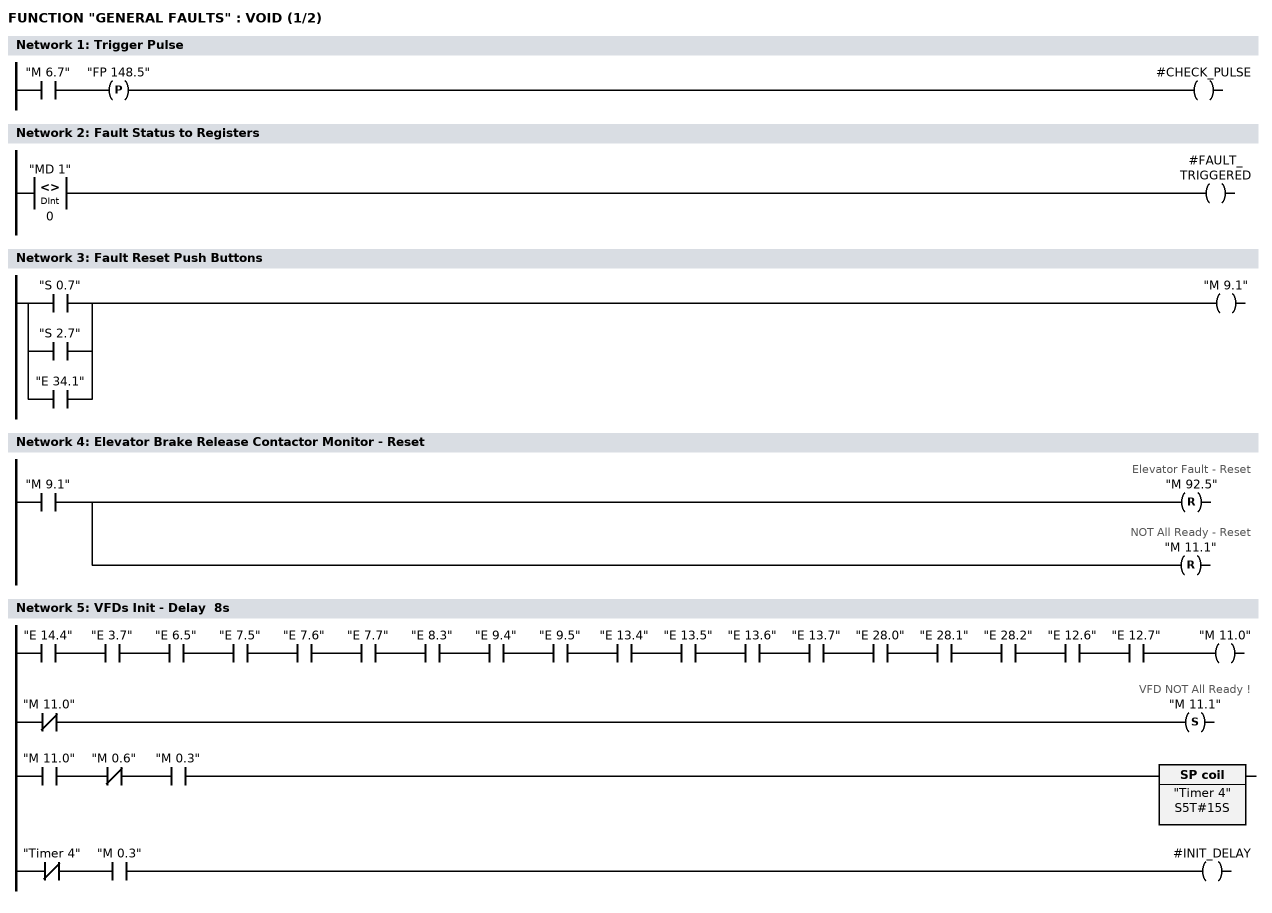

      A     "M 6.7";
      FP    "FP 148.5";
      =     #CHECK_PULSE;
NETWORK
TITLE =Fault Status to Registers

      A(    ;
      L     "MD 1";
      L     0;
      <>D   ;
      )     ;
      =     #FAULT_TRIGGERED;
NETWORK
TITLE =Fault Reset Push Buttons

      A(    ;
      O     "S 0.7";
      O     "S 2.7";
      O     "E 34.1";
      )     ;
      =     "M 9.1";
NETWORK
TITLE =Elevator Brake Release Contactor Monitor - Reset

      A     "M 9.1";
      R     "M 92.5"; // Elevator Fault - Reset
      R     "M 11.1"; // NOT All Ready - Reset
NETWORK
TITLE =VFDs Init - Delay  8s

      A(    ;
      A     "E 14.4";
      A     "E 3.7";
      A     "E 6.5";
      A     "E 7.5";
      A     "E 7.6";
      A     "E 7.7";
      A     "E 8.3";
      A     "E 9.4";
      A     "E 9.5";
      A     "E 13.4";
      A     "E 13.5";
      A     "E 13.6";
      A     "E 13.7";
      A     "E 28.0";
      A     "E 28.1";
      A     "E 28.2";
      A     "E 12.6";
      A     "E 12.7";
      )     ;
      =     "M 11.0";
//;
      AN    "M 11.0";
      S     "M 11.1"; // VFD NOT All Ready !
//;

      A     "M 11.0";
      AN    "M 0.6";
      A     "M 0.3";
      L     S5T#15S;
      SP    "Timer 4";
//;
      AN    "Timer 4";
      A     "M 0.3";
      =     #INIT_DELAY;
NETWORK
TITLE =Motor Temp Control - Fault Check
